(* IEC 61131-3 sources: daoli-st-library/DL_Process (part 13) *)

(* ---- FC_DL_GrateCoolerAirBalanceCalc.st ---- *)
(*
  Name: FC_DL_GrateCoolerAirBalanceCalc
  Category: DL_Process
  Version: 1.0.0
  Round: R91 / 2026-11-25
  开源溯源：clean-room 自研（族 水泥窑篦冷机与预热器，ST 开源生态实测 0 命中，无外部代码引入）
  功能：1) 篦冷机风量收支：把各风室冷却风量逐室求和得总冷却风量 fTotalAirNm3h，
           与窑头抽风（二次风 + 三次风 + 余风）合计 fDraftNm3h 做差，
           差值为正即「多余风量」（须经余风排放），差值为负即「亏缺风量」（抽风大于鼓风）。
        2) 不平衡率 fImbalancePct = |鼓风 − 抽风| / 鼓风 * 100，分母取鼓风侧（可测且恒正），
           方向固定不可交换；该值用于判断风量平衡是否在工艺允许带内。
        3) 平衡判据 fImbalancePct <= fBalMaxPct 输出 xBalanced，供上层选择「投自动调节」或「报警」。
  边界条件：1) 非有限值闸：九路实值入参先过 NOT(x > -DL_BIG AND x < DL_BIG)，同时拦 NaN 与 Inf，
           命中即闸断实值通路（全部输出强制 0.0），不得只置标志（R19）。
        2) 分母零闸：总冷却风量 |fTotalAirNm3h| <= DL_EPS 时不做除法，全部输出清零并判无效。
        3) 物理域闸：任一风室风量或抽风量为负即判无效（负风量属传感器反向或接线错误），
           不取绝对值掩盖符号错误；fBalMaxPct 须落在 (0.0, 100.0] 内，越域视为未组态。
        4) 判据取原始值（R24）：平衡判定使用钳制前的 _fImbalanceRawPct，不得先钳再判。
        5) 物理域钳制：不平衡率钳 0.0 ~ DL_PCT_HI；多余/亏缺风量钳 >= 0（两者互斥，只一支非零）。
        6) 单点赋值（R26）：多余与亏缺由同一差值按符号分支写入，先置 0 再按分支赋值一次，
           不在多处重复写同一变量；纯函数无状态，不做迟滞。
  量纲自证：fTotalAirNm3h / fDraftNm3h / fExcessNm3h / fDeficitNm3h 均为标态体积流量 [Nm3/h]，
           求和与求差两侧同量纲；
           fImbalancePct = |(Nm3/h) − (Nm3/h)| / (Nm3/h) * 100 = 无因次百分数 [%]，量纲合法。
  修订历史 Revision :
    2026-11-25  v1.0.0  R91 首版
*)

FUNCTION FC_DL_GrateCoolerAirBalanceCalc : BOOL
VAR_INPUT
    fChamber1Nm3h    : REAL;   // 1 风室冷却风量 [Nm3/h] / Chamber 1 cooling air flow [Nm3/h]
    fChamber2Nm3h    : REAL;   // 2 风室冷却风量 [Nm3/h] / Chamber 2 cooling air flow [Nm3/h]
    fChamber3Nm3h    : REAL;   // 3 风室冷却风量 [Nm3/h] / Chamber 3 cooling air flow [Nm3/h]
    fChamber4Nm3h    : REAL;   // 4 风室冷却风量 [Nm3/h] / Chamber 4 cooling air flow [Nm3/h]
    fChamber5Nm3h    : REAL;   // 5 风室冷却风量 [Nm3/h] / Chamber 5 cooling air flow [Nm3/h]
    fChamber6Nm3h    : REAL;   // 6 风室冷却风量 [Nm3/h] / Chamber 6 cooling air flow [Nm3/h]
    fDraftNm3h       : REAL;   // 窑头抽风合计（二次+三次+余风）[Nm3/h] / Total kiln-head draft [Nm3/h]
    fBalMaxPct       : REAL;   // 风量平衡允许不平衡率 [%] / Permitted imbalance ratio [%]
END_VAR
VAR_OUTPUT
    fTotalAirNm3h    : REAL;   // 各风室冷却风量合计 [Nm3/h] / Total cooling air flow [Nm3/h]
    fExcessNm3h      : REAL;   // 多余风量（鼓风大于抽风）[Nm3/h] / Excess air flow, blow over draft [Nm3/h]
    fDeficitNm3h     : REAL;   // 亏缺风量（抽风大于鼓风）[Nm3/h] / Deficit air flow, draft over blow [Nm3/h]
    fImbalancePct    : REAL;   // 风量不平衡率 [%] / Air balance imbalance ratio [%]
    xBalanced        : BOOL;   // 风量在允许带内 [bool] / Air balance within tolerance [bool]
    xValid           : BOOL;   // 计算有效标志 [bool] / Calculation valid flag [bool]
END_VAR
VAR
    _fDiffNm3h       : REAL;   // 鼓风减抽风的有符号差值 [Nm3/h] / Signed difference, blow minus draft [Nm3/h]
    _fImbalanceRawPct : REAL;  // 钳制前的不平衡率 [%] / Raw imbalance ratio before limiting [%]
END_VAR
VAR CONSTANT
    DL_EPS           : REAL := 1.0E-9;    // 数值零闸阈值 [-] / Numeric zero gate threshold [-]
    DL_BIG           : REAL := 1.0E12;    // 非有限值闸量级上限 [-] / Finiteness gate magnitude [-]
    DL_PCT           : REAL := 100.0;     // 百分比换算因子 [%] / Percent conversion factor [%]
    DL_PCT_HI        : REAL := 100.0;     // 不平衡率物理上限 [%] / Imbalance physical upper bound [%]
    DL_ZERO_NM3H     : REAL := 0.0;       // 风量零基准 [Nm3/h] / Zero flow reference [Nm3/h]
END_VAR

(* —— 段 1：非有限值闸（R19：闸断实值通路） —— *)
IF NOT (fChamber1Nm3h > -DL_BIG AND fChamber1Nm3h < DL_BIG)
   OR NOT (fChamber2Nm3h > -DL_BIG AND fChamber2Nm3h < DL_BIG)
   OR NOT (fChamber3Nm3h > -DL_BIG AND fChamber3Nm3h < DL_BIG)
   OR NOT (fChamber4Nm3h > -DL_BIG AND fChamber4Nm3h < DL_BIG)
   OR NOT (fChamber5Nm3h > -DL_BIG AND fChamber5Nm3h < DL_BIG)
   OR NOT (fChamber6Nm3h > -DL_BIG AND fChamber6Nm3h < DL_BIG)
   OR NOT (fDraftNm3h > -DL_BIG AND fDraftNm3h < DL_BIG)
   OR NOT (fBalMaxPct > -DL_BIG AND fBalMaxPct < DL_BIG) THEN
    fTotalAirNm3h := 0.0;                   // 输出强制 0.0，切断污染源 / Force zero, cut polluted path
    fExcessNm3h := 0.0;                     // 多余风量强制 0.0 / Excess forced to zero
    fDeficitNm3h := 0.0;                    // 亏缺风量强制 0.0 / Deficit forced to zero
    fImbalancePct := 0.0;                   // 不平衡率强制 0.0 / Imbalance forced to zero
    xBalanced := FALSE;                     // 失效侧不得报平衡 / Must not report balanced when invalid
    xValid := FALSE;                        // 有效位清零 / Validity cleared
    FC_DL_GrateCoolerAirBalanceCalc := FALSE;   // 返回码与有效位同源 / Return mirrors validity
    RETURN;                                 // 立即退出 / Immediate exit
END_IF

(* —— 段 2：风量求和（六室逐室相加，加法顺序不影响结果） —— *)
fTotalAirNm3h := fChamber1Nm3h + fChamber2Nm3h + fChamber3Nm3h
                 + fChamber4Nm3h + fChamber5Nm3h + fChamber6Nm3h;                  // 鼓风合计 [Nm3/h]
_fDiffNm3h := fTotalAirNm3h - fDraftNm3h;                                          // 鼓风 − 抽风 [Nm3/h]

(* —— 段 3：分母零闸（不平衡率的分母是鼓风合计） —— *)
IF ABS(fTotalAirNm3h) <= DL_EPS THEN
    fExcessNm3h := 0.0;                     // 无鼓风即无多余 / No blow, no excess
    fDeficitNm3h := 0.0;                    // 无鼓风即无亏缺 / No blow, no deficit
    fImbalancePct := 0.0;                   // 不平衡率不可算 / Imbalance not computable
    xBalanced := FALSE;                     // 判非平衡 / Not balanced
    xValid := FALSE;                        // 判无效 / Invalid
    FC_DL_GrateCoolerAirBalanceCalc := FALSE;   // 返回码同步 / Return synchronised
    RETURN;                                 // 提前退出 / Early exit
END_IF

_fImbalanceRawPct := ABS(_fDiffNm3h) / fTotalAirNm3h * DL_PCT;                    // 原始不平衡率 [%]

(* —— 段 4：判据（取原始值；单点 BOOL 聚合） —— *)
xValid := (fChamber1Nm3h >= DL_ZERO_NM3H)                                         // 各室风量不得为负
          AND (fChamber2Nm3h >= DL_ZERO_NM3H)
          AND (fChamber3Nm3h >= DL_ZERO_NM3H)
          AND (fChamber4Nm3h >= DL_ZERO_NM3H)
          AND (fChamber5Nm3h >= DL_ZERO_NM3H)
          AND (fChamber6Nm3h >= DL_ZERO_NM3H)
          AND (fDraftNm3h >= DL_ZERO_NM3H)                                        // 抽风量不得为负
          AND (fBalMaxPct > DL_EPS)                                               // 允许带必须为正
          AND (fBalMaxPct <= DL_PCT_HI);                                          // 允许带不得超过 100 %
xBalanced := xValid AND (_fImbalanceRawPct <= fBalMaxPct);                         // 在允许带内才算平衡

(* —— 段 5：多余/亏缺单点分支写入（互斥两支，各自只写一次，R26） —— *)
fExcessNm3h := 0.0;                                                               // 先置零，避免上拍残值
fDeficitNm3h := 0.0;                                                              // 先置零，避免上拍残值
IF _fDiffNm3h > DL_EPS THEN
    fExcessNm3h := _fDiffNm3h;                                                    // 鼓风大于抽风：多余 [Nm3/h]
ELSIF _fDiffNm3h < -DL_EPS THEN
    fDeficitNm3h := ABS(_fDiffNm3h);                                               // 抽风大于鼓风：亏缺 [Nm3/h]
END_IF

(* —— 段 6：输出单点写盘（不平衡率钳制到物理域） —— *)
fImbalancePct := LIMIT(0.0, _fImbalanceRawPct, DL_PCT_HI);                         // 不平衡率钳 0..100 [%]
FC_DL_GrateCoolerAirBalanceCalc := xValid;                                         // 返回码：TRUE = 计算可信

END_FUNCTION

(* ---- FC_DL_GrateCoolerBedResistanceCalc.st ---- *)
(*
  Name: FC_DL_GrateCoolerBedResistanceCalc
  Category: DL_Process
  Version: 1.0.0
  Round: R91 / 2026-11-25
  开源溯源：clean-room 自研（族 水泥窑篦冷机与预热器，ST 开源生态实测 0 命中，无外部代码引入）
  功能：1) 篦床料层阻力按「Ergun 型阻力式的粒度无关简化形」计算：压损正比于料层厚度、
           风量平方与料层堆积密度，反比于开孔率的三次方，
           即 dP = fK * H * rho * (Q/A_open)^2 / 2，A_open = A_total * phi，
           其中 fK 为综合阻力系数（含篦板结构与料层孔隙率经验项）。
        2) 输出三条派生量：料层压损 fBedDpKpa、按开孔率的等效穿孔风速 fOpenVelMs、
           以及压损相对上限的负荷率 fDpLoadPct（用于判断是否接近风机能力极限）。
        3) 压损上限 fDpMaxKpa 为设备许可值，超限只置 xValid=FALSE 并给出超限标志 xDpOver，
           数值本身钳到上限内输出，绝不把越限值伪装成合格值。
  边界条件：1) 非有限值闸：七路实值入参先过 NOT(x > -DL_BIG AND x < DL_BIG)，同时拦 NaN 与 Inf，
           命中即闸断实值通路（全部输出强制 0.0），不得只置标志（R19）。
        2) 分母零闸：料层厚度 fBedHeightM、篦床总面积 fGrateAreaM2 必须 > DL_EPS；
           开孔率 fOpenRatio 必须落在 (DL_PHI_EPS, 1.0] 内 —— 开孔率为 0 或大于 1 均属组态错误，
           直接判无效而非钳制，因为开孔率进三次方，钳制会严重扭曲结果。
        3) 判据取原始值（R24）：压损超限判定使用钳制前的 _fDpRawKpa，
           不得先把压损夹到上限再判是否越限（否则判据恒真）。
        4) 物理域钳制：压损钳 0.0 ~ fDpMaxKpa；穿孔风速钳 0.0 ~ DL_VEL_HI_MS；
           负荷率钳 0.0 ~ DL_LOAD_HI_PCT。
        5) 上限自身校验：fDpMaxKpa 必须 > DL_EPS，为负或零视为未组态，判无效。
        6) 纯函数无状态：不做去抖，堵塞判据的持续性与延时由下游监视 FB 承担。
  量纲自证：开孔面积 A_open = (m2)*(无因次) = m2；
           穿孔风速 = (m3/h)/(m2)/(s/h) = (m3/h)/(m2) * (h/s) = m/s；
           压损 = 无因次 * (m) * (kg/m3) * (m/s)^2 = (kg/m3)*(m2/s2)*(m) = kg/(m*s2) = Pa，
           再除 1000 得 kPa，量纲链自洽。
  修订历史 Revision :
    2026-11-25  v1.0.0  R91 首版
*)

FUNCTION FC_DL_GrateCoolerBedResistanceCalc : BOOL
VAR_INPUT
    fCoolingAirNm3h  : REAL;   // 该风室冷却风量 [Nm3/h] / Cooling air flow of the chamber [Nm3/h]
    fBedHeightM      : REAL;   // 篦床上料层厚度 [m] / Clinker bed height on the grate [m]
    fGrateAreaM2     : REAL;   // 该风室篦床有效面积 [m2] / Effective grate area of the chamber [m2]
    fOpenRatio       : REAL;   // 篦板开孔率（0~1 无因次）[-] / Grate open area ratio, dimensionless [-]
    fBulkDensityKgm3 : REAL;   // 料层堆积密度 [kg/m3] / Clinker bulk density [kg/m3]
    fResistCoef      : REAL;   // 综合阻力系数（含孔隙率经验项）[-] / Combined resistance coefficient [-]
    fDpMaxKpa        : REAL;   // 设备许可料层压损上限 [kPa] / Permitted bed pressure drop [kPa]
END_VAR
VAR_OUTPUT
    fBedDpKpa        : REAL;   // 料层压损 [kPa] / Clinker bed pressure drop [kPa]
    fOpenVelMs       : REAL;   // 篦板穿孔风速 [m/s] / Open-area jet velocity [m/s]
    fDpLoadPct       : REAL;   // 压损对上限的负荷率 [%] / Pressure drop load ratio [%]
    xDpOver          : BOOL;   // 压损超限标志（判定用原始值）[bool] / Pressure drop overrun flag [bool]
    xValid           : BOOL;   // 计算有效标志 [bool] / Calculation valid flag [bool]
END_VAR
VAR
    _fOpenAreaM2     : REAL;   // 篦板有效开孔面积 [m2] / Effective open area of the grate [m2]
    _fOpenVelRawMs   : REAL;   // 钳制前的穿孔风速 [m/s] / Raw open-area velocity [m/s]
    _fDpRawKpa       : REAL;   // 钳制前的原始料层压损 [kPa] / Raw bed pressure drop [kPa]
    _fLoadRawPct     : REAL;   // 钳制前的原始负荷率 [%] / Raw load ratio [%]
END_VAR
VAR CONSTANT
    DL_EPS           : REAL := 1.0E-9;    // 数值零闸阈值 [-] / Numeric zero gate threshold [-]
    DL_PHI_EPS       : REAL := 1.0E-6;    // 开孔率下限阈值 [-] / Open-ratio low gate threshold [-]
    DL_BIG           : REAL := 1.0E12;    // 非有限值闸量级上限 [-] / Finiteness gate magnitude [-]
    DL_SEC_PER_H     : REAL := 3600.0;    // 小时到秒的时基折算 [s/h] / Seconds per hour [s/h]
    DL_PA_PER_KPA    : REAL := 1000.0;    // 帕到千帕的折算 [Pa/kPa] / Pascals per kilopascal [Pa/kPa]
    DL_PHI_HI        : REAL := 1.0;       // 开孔率物理上限 [-] / Open-ratio physical upper bound [-]
    DL_VEL_HI_MS     : REAL := 100.0;     // 穿孔风速物理上限 [m/s] / Jet velocity upper bound [m/s]
    DL_PCT           : REAL := 100.0;     // 百分比换算因子 [%] / Percent conversion factor [%]
    DL_LOAD_HI_PCT   : REAL := 100.0;     // 负荷率物理上限 [%] / Load ratio upper bound [%]
END_VAR

(* —— 段 1：非有限值闸（R19：闸断实值通路） —— *)
IF NOT (fCoolingAirNm3h > -DL_BIG AND fCoolingAirNm3h < DL_BIG)
   OR NOT (fBedHeightM > -DL_BIG AND fBedHeightM < DL_BIG)
   OR NOT (fGrateAreaM2 > -DL_BIG AND fGrateAreaM2 < DL_BIG)
   OR NOT (fOpenRatio > -DL_BIG AND fOpenRatio < DL_BIG)
   OR NOT (fBulkDensityKgm3 > -DL_BIG AND fBulkDensityKgm3 < DL_BIG)
   OR NOT (fResistCoef > -DL_BIG AND fResistCoef < DL_BIG)
   OR NOT (fDpMaxKpa > -DL_BIG AND fDpMaxKpa < DL_BIG) THEN
    fBedDpKpa := 0.0;                       // 输出强制 0.0，切断污染源 / Force zero, cut polluted path
    fOpenVelMs := 0.0;                      // 风速同样强制 0.0 / Velocity forced to zero
    fDpLoadPct := 0.0;                      // 负荷率强制 0.0 / Load ratio forced to zero
    xDpOver := FALSE;                       // 超限位不得在失效时置真 / Overrun must stay false when invalid
    xValid := FALSE;                        // 有效位清零 / Validity cleared
    FC_DL_GrateCoolerBedResistanceCalc := FALSE;   // 返回码与有效位同源 / Return mirrors validity
    RETURN;                                 // 立即退出 / Immediate exit
END_IF

(* —— 段 2：几何与组态域闸（开孔率进三次方，越域一律判无效而非钳制） —— *)
IF (fGrateAreaM2 <= DL_EPS)                                       // 篦床面积不可为零
   OR (fBedHeightM <= DL_EPS)                                     // 料层厚度不可为零
   OR (fOpenRatio <= DL_PHI_EPS)                                  // 开孔率不可为零
   OR (fOpenRatio > DL_PHI_HI)                                    // 开孔率不得大于 1
   OR (fDpMaxKpa <= DL_EPS) THEN                                  // 压损上限必须已组态
    fBedDpKpa := 0.0;                       // 几何不可用即无压损 / No geometry, no drop
    fOpenVelMs := 0.0;                      // 风速不可算 / Velocity not computable
    fDpLoadPct := 0.0;                      // 负荷率不可算 / Load ratio not computable
    xDpOver := FALSE;                       // 失效侧超限位保持假 / Overrun stays false
    xValid := FALSE;                        // 判无效 / Invalid
    FC_DL_GrateCoolerBedResistanceCalc := FALSE;   // 返回码同步 / Return synchronised
    RETURN;                                 // 提前退出 / Early exit
END_IF

(* —— 段 3：主算式（不钳制，先出原始值供段 4 判据使用，R24） —— *)
_fOpenAreaM2 := fGrateAreaM2 * fOpenRatio;                                        // 有效开孔面积 [m2]
_fOpenVelRawMs := fCoolingAirNm3h / _fOpenAreaM2 / DL_SEC_PER_H;                  // 穿孔风速 [m/s]
_fDpRawKpa := fResistCoef * fBedHeightM * fBulkDensityKgm3
              * _fOpenVelRawMs * _fOpenVelRawMs / DL_PA_PER_KPA;                  // 动压式压损 [kPa]
_fLoadRawPct := _fDpRawKpa / fDpMaxKpa * DL_PCT;                                  // 原始负荷率 [%]

(* —— 段 4：判据（全部取原始值；单点 BOOL 聚合避免多处赋 FALSE 覆盖） —— *)
xDpOver := (_fDpRawKpa > fDpMaxKpa);                                              // 压损越上限
xValid := (fCoolingAirNm3h >= 0.0)                                                // 风量不得为负
          AND (fBedHeightM >= 0.0)                                                // 料层厚度不得为负
          AND (fBulkDensityKgm3 > 0.0)                                            // 堆积密度必须为正
          AND (fResistCoef > 0.0)                                                 // 阻力系数必须为正
          AND (_fOpenVelRawMs >= 0.0)                                             // 风速不得为负
          AND (_fDpRawKpa >= 0.0);                                                // 压损不得为负（负压损属符号错误）

(* —— 段 5：输出单点写盘（钳制到物理域内，判定结果已在段 4 定案） —— *)
fBedDpKpa := LIMIT(0.0, _fDpRawKpa, fDpMaxKpa);                                   // 压损钳 0..上限 [kPa]
fOpenVelMs := LIMIT(0.0, _fOpenVelRawMs, DL_VEL_HI_MS);                           // 风速钳 0..上限 [m/s]
fDpLoadPct := LIMIT(0.0, _fLoadRawPct, DL_LOAD_HI_PCT);                           // 负荷率钳 0..100 [%]
FC_DL_GrateCoolerBedResistanceCalc := xValid;                                     // 返回码：TRUE = 计算可信

END_FUNCTION

(* ---- FC_DL_GrateCoolerClinkerTempCalc.st ---- *)
(*
  Name: FC_DL_GrateCoolerClinkerTempCalc
  Category: DL_Process
  Version: 1.0.0
  Round: R91 / 2026-11-25
  开源溯源：clean-room 自研（族 水泥窑篦冷机与预热器，ST 开源生态实测 0 命中，无外部代码引入）
  功能：1) 出篦冷机熟料温度按「熟料放热 = 空气吸热」的稳态能量平衡求解：
           熟料放热 = m_cli * cp_cli * (T_in − T_out)，空气吸热 = m_cli * ratio * cp_air * (T_airOut − T_airIn)，
           两式相等并引入换热效率 eff 后反解出口温度：
           T_out = T_in − eff * ratio * (cp_air / cp_cli) * (T_airOut − T_airIn)。
        2) 输出熟料降温幅度 fCoolDropK，即 T_in − T_out，用于判断冷却能力是否达标。
        3) 温度下限保护：反解结果不得低于 DL_TEMP_LO（环境温度下限），低于即判无效，
           因为能量平衡模型在该区间外已不成立（潜热与辐射项未建模）。
  边界条件：1) 非有限值闸：七路实值入参先过 NOT(x > -DL_BIG AND x < DL_BIG)，同时拦 NaN 与 Inf，
           命中即闸断实值通路（全部输出强制 0.0），不得只置标志（R19）。
        2) 分母零闸：熟料比热 fClinkerCpKjKgK 与风料比 fAirClinkerRatio 均须 > DL_EPS，
           否则反解式分母为零、结果发散，直接判无效。
        3) 参数域闸：换热效率 fEffRatio 必须落在 (0.0, 1.0] 内（效率大于 1 违反热力学第一定律），
           越域视为组态错误判无效，不钳制（钳制会把非法组态伪装成合法）。
        4) 温差方向闸：空气出口温度必须高于空气入口温度，否则无吸热过程，判无效。
        5) 温度下限：反解出口温度 < DL_TEMP_LO 判无效；上限 DL_TEMP_HI 越限判无效。
        6) 判据取原始值（R24）：温度越域判定使用原始反解值 _fOutRawC，钳制只作用于输出量。
  量纲自证：ratio 为风料质量比 [kg/kg] 无因次；cp_air / cp_cli = (kJ/(kg*K))/(kJ/(kg*K)) 无因次；
           eff 无因次；故 eff*ratio*(cp_air/cp_cli)*(T_airOut−T_airIn) 的量纲为 (K)，
           与 T_in [degC] 相减合法（温差以 K 计、绝对温度以 degC 计，差值同尺度）。
  修订历史 Revision :
    2026-11-25  v1.0.0  R91 首版
*)

FUNCTION FC_DL_GrateCoolerClinkerTempCalc : BOOL
VAR_INPUT
    fClinkerInC      : REAL;   // 入篦冷机熟料温度 [degC] / Clinker inlet temperature [degC]
    fAirInC          : REAL;   // 冷却风入口温度（环境）[degC] / Cooling air inlet temperature [degC]
    fAirOutC         : REAL;   // 冷却风出口温度（窑头抽风）[degC] / Cooling air outlet temperature [degC]
    fAirClinkerRatio : REAL;   // 风料质量比 [kg/kg] / Air to clinker mass ratio [kg/kg]
    fAirCpKjKgK      : REAL;   // 空气定压比热 [kJ/(kg*K)] / Air specific heat at constant pressure [kJ/(kg*K)]
    fClinkerCpKjKgK  : REAL;   // 熟料比热 [kJ/(kg*K)] / Clinker specific heat [kJ/(kg*K)]
    fEffRatio        : REAL;   // 篦床换热效率（0~1 无因次）[-] / Grate heat exchange efficiency, dimensionless [-]
END_VAR
VAR_OUTPUT
    fClinkerOutC     : REAL;   // 出篦冷机熟料温度 [degC] / Clinker outlet temperature [degC]
    fCoolDropK       : REAL;   // 熟料降温幅度 [K] / Clinker temperature drop [K]
    xTempLow         : BOOL;   // 出口温度低于下限标志 [bool] / Outlet below lower bound flag [bool]
    xValid           : BOOL;   // 计算有效标志 [bool] / Calculation valid flag [bool]
END_VAR
VAR
    _fCpRatio        : REAL;   // 空气与熟料比热之比 [-] / Ratio of air to clinker specific heat [-]
    _fAirDeltaK      : REAL;   // 空气温升 [K] / Air temperature rise [K]
    _fOutRawC        : REAL;   // 钳制前的原始出口温度 [degC] / Raw outlet temperature before limiting [degC]
    _fDropRawK       : REAL;   // 钳制前的原始降温幅度 [K] / Raw temperature drop before limiting [K]
END_VAR
VAR CONSTANT
    DL_EPS           : REAL := 1.0E-9;    // 数值零闸阈值 [-] / Numeric zero gate threshold [-]
    DL_BIG           : REAL := 1.0E12;    // 非有限值闸量级上限 [-] / Finiteness gate magnitude [-]
    DL_TEMP_LO       : REAL := -50.0;     // 熟料出口温度物理下限 [degC] / Clinker outlet lower bound [degC]
    DL_TEMP_HI       : REAL := 400.0;     // 熟料出口温度物理上限 [degC] / Clinker outlet upper bound [degC]
    DL_EFF_HI        : REAL := 1.0;       // 换热效率物理上限（热力学第一定律）[-] / Efficiency upper bound [-]
    DL_ZERO_K        : REAL := 0.0;       // 温差零基准 [K] / Zero temperature-difference reference [K]
END_VAR

(* —— 段 1：非有限值闸（R19：闸断实值通路） —— *)
IF NOT (fClinkerInC > -DL_BIG AND fClinkerInC < DL_BIG)
   OR NOT (fAirInC > -DL_BIG AND fAirInC < DL_BIG)
   OR NOT (fAirOutC > -DL_BIG AND fAirOutC < DL_BIG)
   OR NOT (fAirClinkerRatio > -DL_BIG AND fAirClinkerRatio < DL_BIG)
   OR NOT (fAirCpKjKgK > -DL_BIG AND fAirCpKjKgK < DL_BIG)
   OR NOT (fClinkerCpKjKgK > -DL_BIG AND fClinkerCpKjKgK < DL_BIG)
   OR NOT (fEffRatio > -DL_BIG AND fEffRatio < DL_BIG) THEN
    fClinkerOutC := 0.0;                    // 输出强制 0.0，切断污染源 / Force zero, cut polluted path
    fCoolDropK := 0.0;                      // 降温幅度强制 0.0 / Drop forced to zero
    xTempLow := FALSE;                      // 失效侧不得报低温 / Must not report low temp when invalid
    xValid := FALSE;                        // 有效位清零 / Validity cleared
    FC_DL_GrateCoolerClinkerTempCalc := FALSE;   // 返回码与有效位同源 / Return mirrors validity
    RETURN;                                 // 立即退出 / Immediate exit
END_IF

(* —— 段 2：分母零闸与参数域闸（比热、风料比为零则反解发散） —— *)
IF (fClinkerCpKjKgK <= DL_EPS)                                    // 熟料比热不可为零
   OR (fAirClinkerRatio <= DL_EPS)                                // 风料比不可为零
   OR (fAirCpKjKgK <= DL_EPS)                                     // 空气比热不可为零
   OR (fEffRatio <= DL_EPS)                                       // 换热效率不可为零
   OR (fEffRatio > DL_EFF_HI) THEN                                // 换热效率不得大于 1（热力学第一定律）
    fClinkerOutC := 0.0;                    // 参数不可用即无出口温度 / No parameter, no outlet temperature
    fCoolDropK := 0.0;                      // 降温幅度不可算 / Drop not computable
    xTempLow := FALSE;                      // 失效侧低温位保持假 / Low-temp flag stays false
    xValid := FALSE;                        // 判无效 / Invalid
    FC_DL_GrateCoolerClinkerTempCalc := FALSE;   // 返回码同步 / Return synchronised
    RETURN;                                 // 提前退出 / Early exit
END_IF

(* —— 段 3：主算式（不钳制，先出原始值供段 4 判据使用，R24） —— *)
_fCpRatio := fAirCpKjKgK / fClinkerCpKjKgK;                                       // 比热之比 [-]
_fAirDeltaK := fAirOutC - fAirInC;                                                // 空气温升 [K]
_fOutRawC := fClinkerInC - fEffRatio * fAirClinkerRatio * _fCpRatio * _fAirDeltaK; // 出口温度反解 [degC]
_fDropRawK := fClinkerInC - _fOutRawC;                                            // 降温幅度 [K]

(* —— 段 4：判据（取原始值；单点 BOOL 聚合避免多处赋 FALSE 覆盖） —— *)
xTempLow := (_fOutRawC < DL_TEMP_LO);                                             // 出口低于物理下限
xValid := (_fAirDeltaK > DL_ZERO_K)                                               // 空气必须吸热（出口高于入口）
          AND (_fOutRawC >= DL_TEMP_LO)                                           // 不跌破物理下限
          AND (_fOutRawC <= DL_TEMP_HI)                                           // 不超出物理上限
          AND (_fDropRawK >= DL_ZERO_K)                                           // 降温幅度不得为负（方向固定）
          AND (fClinkerInC > DL_TEMP_LO);                                         // 入口温度本身须在物理域内

(* —— 段 5：输出单点写盘（钳制到物理域内，判定结果已在段 4 定案） —— *)
fClinkerOutC := LIMIT(DL_TEMP_LO, _fOutRawC, DL_TEMP_HI);                          // 出口温度钳物理域 [degC]
fCoolDropK := MAX(DL_ZERO_K, _fDropRawK);                                          // 降温幅度钳 >= 0 [K]
FC_DL_GrateCoolerClinkerTempCalc := xValid;                                        // 返回码：TRUE = 计算可信

END_FUNCTION

(* ---- FC_DL_GrateCoolerHeatRecoveryCalc.st ---- *)
(*
  Name: FC_DL_GrateCoolerHeatRecoveryCalc
  Category: DL_Process
  Version: 1.0.0
  Round: R91 / 2026-11-25
  开源溯源：clean-room 自研（族 水泥窑篦冷机与预热器，ST 开源生态实测 0 命中，无外部代码引入）
  功能：1) 回收热量取「二次风显热 + 三次风显热」，两者均以环境温度为基准，风侧按定压比热折算，
           即 fRecoveredHeatKw = (V2*cp*(T2-Tamb) + V3*cp*(T3-Tamb)) / 3600，单位 kW，
           3600 为 kJ/h 到 kW 的时基折算系数。
        2) 熟料可供显热取「熟料量 × 熟料比热 × (入篦床温度 − 出篦床温度)」，
           即 fClinkerHeatKw = m*1000*cpCli*(Tin-Tout) / 3600，单位 kW，
           1000 为 t 到 kg 的质量折算系数；该项是回收率的物理分母（可供热上限）。
        3) 热回收率 fRecoveryPct = 回收热量 / 熟料可供显热 * 100，钳制 0.0 ~ 100.0 %，
           回收率超过 100 % 在物理上不可能，判为测量链路故障而非效率优异。
  边界条件：1) 非有限值闸：九路实值入参先过 NOT(x > -DL_BIG AND x < DL_BIG)，该式同时拦 NaN 与 Inf，
           命中即闸断实值通路（全部输出强制 0.0），不得只置 xValid 而把 NaN 传给下游（R19）。
        2) 分母零闸：风侧比热 fAirCpKjNm3K 与熟料比热 fClinkerCp 均须 > DL_EPS，
           熟料可供显热 |fClinkerHeatKw| > DL_EPS 才允许做除法，否则判无效并清零。
        3) 判据取原始值（R24）：回收率越限判定使用 LIMIT 之前的原始值 _fRecoveryRawPct，
           不得先把回收率夹到 0~100 再判超域（否则判据恒真，域闸静默失效）。
        4) 物理域钳制：回收率钳 0.0 ~ 100.0 %；两路风量与熟料量不得为负（负值即传感器反向，判无效）。
        5) 温度方向校验：二次/三次风温低于环境温度、或熟料出口温度高于入口温度，均属非冷却工况，
           判无效而不取绝对值掩盖符号错误。
        6) 纯函数无状态：本件不做迟滞与去抖，滤波与报警延时由下游监视 FB 承担。
  量纲自证：fRecoveredHeatKw = (Nm3/h)*(kJ/(Nm3*K))*(K) / (s/h) = (kJ/h)/(s/h) = kJ/s = kW；
           fClinkerHeatKw   = (t/h)*(kg/t)*(kJ/(kg*K))*(K) / (s/h) = (kJ/h)/(s/h) = kW；
           fRecoveryPct     = (kW)/(kW)*100 = 无因次百分数 [%]，比量两侧同量纲，量纲关系合法。
  修订历史 Revision :
    2026-11-25  v1.0.0  R91 首版
*)

FUNCTION FC_DL_GrateCoolerHeatRecoveryCalc : BOOL
VAR_INPUT
    fSecAirNm3h      : REAL;   // 二次风标态体积流量 [Nm3/h] / Secondary air normal flow [Nm3/h]
    fTerAirNm3h      : REAL;   // 三次风标态体积流量 [Nm3/h] / Tertiary air normal flow [Nm3/h]
    fSecAirTempC     : REAL;   // 二次风温度 [degC] / Secondary air temperature [degC]
    fTerAirTempC     : REAL;   // 三次风温度 [degC] / Tertiary air temperature [degC]
    fAmbientC        : REAL;   // 环境基准温度 [degC] / Ambient reference temperature [degC]
    fClinkerTph      : REAL;   // 熟料产量 [t/h] / Clinker production rate [t/h]
    fClinkerInC      : REAL;   // 入篦床熟料温度 [degC] / Clinker inlet temperature [degC]
    fClinkerOutC     : REAL;   // 出篦床熟料温度 [degC] / Clinker outlet temperature [degC]
    fAirCpKjNm3K     : REAL;   // 风侧定压比热 [kJ/(Nm3*K)] / Air specific heat at constant pressure [kJ/(Nm3*K)]
    fClinkerCpKjKgK  : REAL;   // 熟料比热 [kJ/(kg*K)] / Clinker specific heat [kJ/(kg*K)]
END_VAR
VAR_OUTPUT
    fRecoveredHeatKw : REAL;   // 二次+三次风回收热量 [kW] / Recovered heat by secondary and tertiary air [kW]
    fClinkerHeatKw   : REAL;   // 熟料可供显热 [kW] / Clinker available sensible heat [kW]
    fRecoveryPct     : REAL;   // 热回收率 [%] / Heat recovery ratio [%]
    xValid           : BOOL;   // 计算有效标志 [bool] / Calculation valid flag [bool]
END_VAR
VAR
    _fSecHeatKjh     : REAL;   // 二次风显热 [kJ/h] / Secondary air sensible heat [kJ/h]
    _fTerHeatKjh     : REAL;   // 三次风显热 [kJ/h] / Tertiary air sensible heat [kJ/h]
    _fRecoveredKjh   : REAL;   // 回收热量合计（钳制前）[kJ/h] / Total recovered heat before limiting [kJ/h]
    _fClinkerKjh     : REAL;   // 熟料可供显热（钳制前）[kJ/h] / Clinker sensible heat before limiting [kJ/h]
    _fRecoveryRawPct : REAL;   // 钳制前的原始回收率 [%] / Raw recovery before limiting [%]
END_VAR
VAR CONSTANT
    DL_EPS           : REAL := 1.0E-9;    // 数值零闸阈值 [-] / Numeric zero gate threshold [-]
    DL_BIG           : REAL := 1.0E12;    // 非有限值闸量级上限 [-] / Finiteness gate magnitude [-]
    DL_SEC_PER_H     : REAL := 3600.0;    // 小时到秒的时基折算 [s/h] / Seconds per hour [s/h]
    DL_KG_PER_T      : REAL := 1000.0;    // 吨到千克的质量折算 [kg/t] / Kilograms per tonne [kg/t]
    DL_PCT           : REAL := 100.0;     // 百分比换算因子 [%] / Percent conversion factor [%]
    DL_REC_LO_PCT    : REAL := 0.0;       // 回收率物理域下限 [%] / Recovery physical domain low [%]
    DL_REC_HI_PCT    : REAL := 100.0;     // 回收率物理域上限 [%] / Recovery physical domain high [%]
END_VAR

(* —— 段 1：非有限值闸（R19：闸断实值通路，NaN/Inf 一律不得流到输出） —— *)
IF NOT (fSecAirNm3h > -DL_BIG AND fSecAirNm3h < DL_BIG)
   OR NOT (fTerAirNm3h > -DL_BIG AND fTerAirNm3h < DL_BIG)
   OR NOT (fSecAirTempC > -DL_BIG AND fSecAirTempC < DL_BIG)
   OR NOT (fTerAirTempC > -DL_BIG AND fTerAirTempC < DL_BIG)
   OR NOT (fAmbientC > -DL_BIG AND fAmbientC < DL_BIG)
   OR NOT (fClinkerTph > -DL_BIG AND fClinkerTph < DL_BIG)
   OR NOT (fClinkerInC > -DL_BIG AND fClinkerInC < DL_BIG)
   OR NOT (fClinkerOutC > -DL_BIG AND fClinkerOutC < DL_BIG)
   OR NOT (fAirCpKjNm3K > -DL_BIG AND fAirCpKjNm3K < DL_BIG)
   OR NOT (fClinkerCpKjKgK > -DL_BIG AND fClinkerCpKjKgK < DL_BIG) THEN
    fRecoveredHeatKw := 0.0;                // 输出强制 0.0，切断污染源 / Force zero, cut polluted path
    fClinkerHeatKw := 0.0;                  // 熟料显热同样强制 0.0 / Clinker heat forced to zero
    fRecoveryPct := 0.0;                    // 回收率强制 0.0 / Recovery forced to zero
    xValid := FALSE;                        // 有效位清零 / Validity cleared
    FC_DL_GrateCoolerHeatRecoveryCalc := FALSE;   // 返回码与有效位同源 / Return mirrors validity
    RETURN;                                 // 立即退出 / Immediate exit
END_IF

(* —— 段 2：比热零闸（R4：除法前先过零闸，且闸的是分母本身） —— *)
IF ABS(fAirCpKjNm3K) <= DL_EPS OR ABS(fClinkerCpKjKgK) <= DL_EPS THEN
    fRecoveredHeatKw := 0.0;                // 比热缺失即无法折算 / No specific heat, no conversion
    fClinkerHeatKw := 0.0;                  // 熟料显热不可算 / Clinker heat not computable
    fRecoveryPct := 0.0;                    // 回收率不可算 / Recovery not computable
    xValid := FALSE;                        // 判无效 / Invalid
    FC_DL_GrateCoolerHeatRecoveryCalc := FALSE;   // 返回码同步 / Return synchronised
    RETURN;                                 // 提前退出 / Early exit
END_IF

(* —— 段 3：主算式（不做任何钳制，先出原始值供段 4 判据使用，R24） —— *)
_fSecHeatKjh := fSecAirNm3h * fAirCpKjNm3K * (fSecAirTempC - fAmbientC);          // 二次风显热 [kJ/h]
_fTerHeatKjh := fTerAirNm3h * fAirCpKjNm3K * (fTerAirTempC - fAmbientC);          // 三次风显热 [kJ/h]
_fRecoveredKjh := _fSecHeatKjh + _fTerHeatKjh;                                    // 回收热量合计 [kJ/h]
_fClinkerKjh := fClinkerTph * DL_KG_PER_T * fClinkerCpKjKgK
                * (fClinkerInC - fClinkerOutC);                                   // 熟料可供显热 [kJ/h]

(* —— 段 4：分母零闸（熟料可供显热为回收率的分母） —— *)
IF ABS(_fClinkerKjh) <= DL_EPS THEN
    fRecoveredHeatKw := 0.0;                // 无可供热即无回收率 / No source heat, no recovery
    fClinkerHeatKw := 0.0;                  // 分母侧同步清零 / Denominator side zeroed
    fRecoveryPct := 0.0;                    // 回收率清零 / Recovery zeroed
    xValid := FALSE;                        // 判无效 / Invalid
    FC_DL_GrateCoolerHeatRecoveryCalc := FALSE;   // 返回码同步 / Return synchronised
    RETURN;                                 // 提前退出 / Early exit
END_IF

_fRecoveryRawPct := _fRecoveredKjh / _fClinkerKjh * DL_PCT;                       // 原始回收率 [%]

(* —— 段 5：物理域与符号校验（判据全部取原始值，单点 BOOL 聚合避免多处赋 FALSE 覆盖） —— *)
xValid := (fSecAirNm3h >= 0.0)                                        // 二次风量不得为负
          AND (fTerAirNm3h >= 0.0)                                    // 三次风量不得为负
          AND (fClinkerTph >= 0.0)                                    // 熟料量不得为负
          AND (_fRecoveredKjh >= 0.0)                                 // 风温低于环境温度属非回收工况
          AND (_fClinkerKjh > 0.0)                                    // 熟料出口必须低于入口
          AND (_fRecoveryRawPct >= DL_REC_LO_PCT)                     // 不低于物理域下限
          AND (_fRecoveryRawPct <= DL_REC_HI_PCT);                    // 不高于物理域上限（>100 % 物理不可能）

(* —— 段 6：输出单点写盘（数值钳制到物理域内，有效位已在段 5 定案） —— *)
fRecoveredHeatKw := _fRecoveredKjh / DL_SEC_PER_H;                                        // 折算为 kW
fClinkerHeatKw := _fClinkerKjh / DL_SEC_PER_H;                                            // 折算为 kW
fRecoveryPct := LIMIT(DL_REC_LO_PCT, _fRecoveryRawPct, DL_REC_HI_PCT);                    // 回收率钳 0..100 [%]
FC_DL_GrateCoolerHeatRecoveryCalc := xValid;                                              // 返回码：TRUE = 计算可信

END_FUNCTION

(* ---- FC_DL_GreenSandCompactabilityCalc.st ---- *)
(*
 * FC_DL_GreenSandCompactabilityCalc | C1 | DL_Process
 * 功能：由含水量反算紧实率并判定是否落在工艺带       单位：水分 [%]、紧实率 [%]、系数 [%/%、1]
 * 工况边界：w = a + b×CB 的反解 CB = (w−a)/b，b 须 >0（本件强制 b≠0，否则判 9714）；工艺带 30~45 %（含端点，浮点比较用容差）；a、b 与水分须有限
 * 代数值回代：w=3.0 %、a=1.2、b=0.04 → CB=(3.0−1.2)/0.04=45 %，落在 30~45 → xInRange=TRUE（与 spec 回代行一致）
 * 开源溯源：clean-room 自研，未复制任何第三方代码（无外部来源）
 *)
FUNCTION FC_DL_GreenSandCompactabilityCalc : BOOL
VAR_INPUT
    rMoisturePct : REAL := 3.0;      // 型砂含水量 | green sand moisture [%]
    rA           : REAL := 1.2;      // 经验式截距 | empirical intercept [%]
    rB           : REAL := 0.04;     // 经验式斜率 | empirical slope [%/%]
END_VAR
VAR_OUTPUT
    rCompactabilityPct : REAL;       // 紧实率 | compactability [%]
    xInRange           : BOOL;       // 落在工艺带 30~45 | inside the process band 30 to 45
    xValid             : BOOL;       // 输出有效 | outputs valid
    nFaultCode         : INT;        // 0=无 / 9714=斜率或水分非法 | 0 none, 9714 illegal slope or moisture
END_VAR
VAR
    xFinW : BOOL;                    // 水分有限性 | moisture is finite
    xFinA : BOOL;                    // 截距有限性 | intercept is finite
    xFinB : BOOL;                    // 斜率有限性 | slope is finite
END_VAR
VAR CONSTANT
    DL_GSC_LO  : REAL := 30.0;       // 工艺带下限 | process band lower bound [%]
    DL_GSC_HI  : REAL := 45.0;       // 工艺带上限 | process band upper bound [%]
    DL_GSC_EPS : REAL := 1.0E-6;     // 浮点比较容差 | floating comparison tolerance [%]
    DL_GSC_BMIN: REAL := 1.0E-9;     // 斜率下限（防零除）| slope lower bound guarding the division [%/%]
END_VAR

// 段1｜非有限闸（R19）
xFinW := (rMoisturePct = rMoisturePct) AND ((rMoisturePct - rMoisturePct) = 0.0);
xFinA := (rA = rA) AND ((rA - rA) = 0.0);
xFinB := (rB = rB) AND ((rB - rB) = 0.0);
IF (NOT xFinW) OR (NOT xFinA) OR (NOT xFinB) THEN
    rCompactabilityPct := 0.0;       // 安全值：紧实率 0 | safe value, zero compactability
    xInRange := FALSE;
    xValid := FALSE;
    nFaultCode := 9714;
    FC_DL_GreenSandCompactabilityCalc := FALSE;
    RETURN;
END_IF

// 段2｜域闸：斜率入分母必须为正，水分不得为负
IF (rB <= DL_GSC_BMIN) OR (rMoisturePct < 0.0) THEN
    rCompactabilityPct := 0.0;
    xInRange := FALSE;
    xValid := FALSE;
    nFaultCode := 9714;
    FC_DL_GreenSandCompactabilityCalc := FALSE;
    RETURN;
END_IF

// 段3｜算法：CB = (w − a)/b
rCompactabilityPct := (rMoisturePct - rA) / rB;

// 段4｜工艺带判定（判据与出口同源于原始水分推算值）
xInRange := (rCompactabilityPct >= (DL_GSC_LO - DL_GSC_EPS))
             AND (rCompactabilityPct <= (DL_GSC_HI + DL_GSC_EPS));
nFaultCode := 0;
xValid := TRUE;
FC_DL_GreenSandCompactabilityCalc := TRUE;
END_FUNCTION

(* ---- FC_DL_GreenSandMoistureTargetCalc.st ---- *)
(*
 * FC_DL_GreenSandMoistureTargetCalc | C2 | DL_Process
 * 功能：由紧实率反算湿型砂水分目标（线性经验式）       单位：紧实率 [%]、水分 [%]、系数 [%/%、1]
 * 工况边界：经验式 w = a + b×CB，a=1.2 %、b=0.04 %/%（spec 采纳值，回代 38 → 2.72 %，落在湿型砂 2.5~3.5 % 合理区间）；紧实率按物理域钳位 [20,60] %，越界置信息位且判据取自未钳位原值；系数 b 须 >0
 * 代数值回代：CB=38 %、a=1.2、b=0.04 → w=1.2+0.04×38=2.72 %（与 spec 采纳回代值一致）
 * 系数修正说明：spec 初版给 a=0.55 / b=0.0525，回代 38 得 2.545 % 偏离湿型砂常规区间，spec 已明确改用 a=1.2 / b=0.04，本件按采纳值实现
 * 开源溯源：clean-room 自研，未复制任何第三方代码（无外部来源）
 *)
FUNCTION FC_DL_GreenSandMoistureTargetCalc : BOOL
VAR_INPUT
    rCompactabilityPct : REAL := 38.0;  // 紧实率 | compactability [%]
    rA                 : REAL := 1.2;   // 经验式截距 | empirical intercept [%]
    rB                 : REAL := 0.04;  // 经验式斜率 | empirical slope [%/%]
END_VAR
VAR_OUTPUT
    rTargetMoisturePct : REAL;          // 目标水分 | target moisture [%]
    rCbUsed            : REAL;          // 实际参与计算的紧实率（已钳位）| compactability actually used, clamped [%]
    xClamped           : BOOL;          // 紧实率越界被钳位（信息级）| compactability clamped, informational
    xValid             : BOOL;          // 输出有效 | outputs valid
END_VAR
VAR
    xFinCb : BOOL;                      // 紧实率有限性 | compactability is finite
    xFinA  : BOOL;                      // 截距有限性 | intercept is finite
    xFinB  : BOOL;                      // 斜率有限性 | slope is finite
END_VAR
VAR CONSTANT
    DL_GSM_CB_LO : REAL := 20.0;        // 紧实率物理下限 | compactability lower bound [%]
    DL_GSM_CB_HI : REAL := 60.0;        // 紧实率物理上限 | compactability upper bound [%]
END_VAR

// 段1｜非有限闸（R19）
xFinCb := (rCompactabilityPct = rCompactabilityPct) AND ((rCompactabilityPct - rCompactabilityPct) = 0.0);
xFinA := (rA = rA) AND ((rA - rA) = 0.0);
xFinB := (rB = rB) AND ((rB - rB) = 0.0);
IF (NOT xFinCb) OR (NOT xFinA) OR (NOT xFinB) THEN
    rTargetMoisturePct := 0.0;          // 安全值：目标水分 0 | safe value, zero target
    rCbUsed := 0.0;
    xClamped := FALSE;
    xValid := FALSE;
    FC_DL_GreenSandMoistureTargetCalc := FALSE;
    RETURN;
END_IF

// 段2｜域闸：斜率必须为正（经验式单调增，否则反算无意义）
IF rB <= 0.0 THEN
    rTargetMoisturePct := 0.0;
    rCbUsed := 0.0;
    xClamped := FALSE;
    xValid := FALSE;
    FC_DL_GreenSandMoistureTargetCalc := FALSE;
    RETURN;
END_IF

// 段3｜域钳位：越界标志取自未钳位原值（R24）
IF rCompactabilityPct < DL_GSM_CB_LO THEN
    xClamped := TRUE;
    rCbUsed := DL_GSM_CB_LO;
ELSIF rCompactabilityPct > DL_GSM_CB_HI THEN
    xClamped := TRUE;
    rCbUsed := DL_GSM_CB_HI;
ELSE
    xClamped := FALSE;
    rCbUsed := rCompactabilityPct;
END_IF

// 段4｜算法：w = a + b×CB
rTargetMoisturePct := rA + rB * rCbUsed;
xValid := TRUE;
FC_DL_GreenSandMoistureTargetCalc := TRUE;
END_FUNCTION

(* ---- FC_DL_GreenStrengthIndexCalc.st ---- *)
(*
  Component : FC_DL_GreenStrengthIndexCalc
  Category  : DL_Process
  Type      : FC
  Complexity: C2
  VERSION   : v1.0.0
  功能      : 生坯强度指数核算：按压制成型压力、润滑剂含量与生坯密度算无量纲强度指数，并与安全阈值比较给出脱模安全判定。
  开源溯源  : 道莅原创 clean-room 自研（无外部代码引用）｜License: MIT
  边界条件  : ① 参考密度与安全阈值须 > 1e-9，压制压力须非负，润滑剂含量须在 0~5 % 内，否则返回哨兵 -1；
              ② 压力项取开方（压力对强度是次线性贡献），开方前已钳位非负；
              ③ 润滑剂含量越高生坯强度越低，折算系数下限钳位 0.3。
*)
FUNCTION FC_DL_GreenStrengthIndexCalc : REAL
VAR_INPUT
    fPressMPa    : REAL;   (* 压制压力 [MPa] Compaction pressure *)
    fLubePct     : REAL;   (* 润滑剂含量 [%] Lubricant content *)
    fGreenDens   : REAL;   (* 生坯密度 [g/cm³] Green density *)
    fDensRef     : REAL;   (* 参考密度（工艺目标） [g/cm³] Reference density *)
    fSafeIdx     : REAL;   (* 脱模安全指数阈值 [-] Safe ejection index threshold *)
END_VAR
VAR_OUTPUT
    fStrengthIdx : REAL;  (* 生坯强度指数 [-] Green strength index *)
    fLubeFactor  : REAL;  (* 润滑剂折减因子 [-] Lubricant reduction factor *)
    xEjectSafe   : BOOL;  (* 脱模安全标志 [-] Safe ejection flag *)
    xValid       : BOOL;  (* 计算有效性标志 [-] Calculation valid flag *)
END_VAR
VAR CONSTANT
    DL_EPS      : REAL := 1.0E-9;   (* 除零判定容差 [无量纲] Divide-by-zero tolerance *)
    DL_PCT_BASE : REAL := 100.0;    (* 百分比基准 [%] Percent base *)
    DL_GAIN     : REAL := 3.0;      (* 压力项标定增益 [-] Pressure term gain *)
    DL_LUBE_K   : REAL := 0.9;      (* 润滑剂折减系数 [-] Lubricant reduction coefficient *)
    DL_LUBE_MAX : REAL := 5.0;      (* 润滑剂含量上限 [%] Lubricant upper bound *)
    DL_LF_MIN   : REAL := 0.3;      (* 润滑剂因子下限 [-] Lubricant factor floor *)
    DL_ZERO     : REAL := 0.0;      (* 零常量 [无量纲] Zero constant *)
END_VAR
VAR
    fPressPos : REAL;   (* 非负压制压力 [MPa] Non-negative pressure *)
END_VAR
(* 出口预置：四出口统一预置 *)
fStrengthIdx := 0.0; fLubeFactor := 1.0; xEjectSafe := FALSE; xValid := FALSE;
(* 非有限拦截：自反判 NaN，自身差值判 Inf *)
IF (fPressMPa <> fPressMPa) OR ((fPressMPa - fPressMPa) <> 0.0)
   OR (fLubePct <> fLubePct) OR ((fLubePct - fLubePct) <> 0.0)
   OR (fGreenDens <> fGreenDens) OR ((fGreenDens - fGreenDens) <> 0.0)
   OR (fDensRef <> fDensRef) OR ((fDensRef - fDensRef) <> 0.0)
   OR (fSafeIdx <> fSafeIdx) OR ((fSafeIdx - fSafeIdx) <> 0.0) THEN
    FC_DL_GreenStrengthIndexCalc := -1.0;  (* 哨兵 -1：输入非有限 / Sentinel -1 non-finite *)
    RETURN;
END_IF
(* 组态域闸：参考密度与安全阈值为比例基，润滑剂含量与压力取可表区间 *)
IF (fDensRef <= DL_EPS) OR (fSafeIdx <= DL_EPS) OR (fPressMPa < DL_ZERO)
   OR (fLubePct < DL_ZERO) OR (fLubePct > DL_LUBE_MAX) OR (fGreenDens < DL_ZERO) THEN
    FC_DL_GreenStrengthIndexCalc := -1.0;  (* 哨兵 -1：组态非法 / Sentinel -1 bad config *)
    RETURN;
END_IF
(* 润滑剂折减因子：含量越高强度越低，下限钳位 0.3 防归零 *)
fLubeFactor := 1.0 - (fLubePct / DL_PCT_BASE) * DL_LUBE_K;
IF fLubeFactor < DL_LF_MIN THEN
    fLubeFactor := DL_LF_MIN;                 (* 下限钳位 [-] / Lower clamp *)
END_IF
(* 压力项非负钳位后开方（开方前判非负） *)
fPressPos := fPressMPa;
IF fPressPos < DL_ZERO THEN
    fPressPos := DL_ZERO;
END_IF
(* 强度指数：sqrt(p) × 增益 × 润滑剂因子 × 密度比，参考密度已过域闸 *)
fStrengthIdx := SQRT(fPressPos) * DL_GAIN * fLubeFactor * (fGreenDens / fDensRef);
(* 脱模安全判定：指数达阈值即可安全脱模 *)
xEjectSafe := fStrengthIdx >= fSafeIdx;
xValid := TRUE;                               (* 链路有效 / Chain valid *)
FC_DL_GreenStrengthIndexCalc := fStrengthIdx; (* 返回强度指数 [-] / Return strength index *)
END_FUNCTION

(* ---- FC_DL_HexChromeTriRatioCalc.st ---- *)
(*
  DL Factory R83 | FC_DL_HexChromeTriRatioCalc
  功能：算六价铬与三价铬浓度比，判定镀液老化并给出需氧化的三价铬过量值。
  开源溯源：无（clean-room 自研，依据公开工艺公式，来源=行业通用公式，许可证=MIT，借鉴点=公式结构）
  规则：R1-R21 全遵守
*)
FUNCTION FC_DL_HexChromeTriRatioCalc : REAL
VAR_INPUT
    fCr6Gpl   : REAL; // 六价铬浓度 [g/L] / Hexavalent chromium concentration [g/L]
    fCr3Gpl   : REAL; // 三价铬浓度 [g/L] / Trivalent chromium concentration [g/L]
    fRatioMin : REAL; // 允许最低六/三比值 [-]/ Minimum allowed hex-to-tri ratio [-]
    fTempC    : REAL; // 槽液温度 [°C] / Bath temperature [degC]
END_VAR
VAR_OUTPUT
    fRatio     : REAL; // 六价/三价比值 [-]/ Hex-to-tri concentration ratio [-]
    fCr3Excess : REAL; // 三价铬过量（需氧化去除量，负值按零）[g/L] / Excess trivalent [g/L]
    xAged      : BOOL; // 老化判定（TRUE=三价累积超限）/ Ageing flag, TRUE = build-up
    xValid     : BOOL; // 计算有效性标志 / Calculation validity flag
END_VAR
VAR
    fCr3Limit : REAL; // 三价铬允许上限 [g/L] / Allowed trivalent ceiling [g/L]
END_VAR
// 出口预置：四出口统一预置，老化标志预置 FALSE（安全侧）
fRatio := 0.0; fCr3Excess := 0.0; xAged := FALSE; xValid := FALSE;
// 非有限拦截 + 量纲自检（R20/R21）
IF NOT (fCr6Gpl > -1.0E30 AND fCr6Gpl < 1.0E30) OR NOT (fCr3Gpl > -1.0E30 AND fCr3Gpl < 1.0E30) OR NOT (fRatioMin > -1.0E30 AND fRatioMin < 1.0E30) OR NOT (fTempC > -1.0E30 AND fTempC < 1.0E30) OR fCr6Gpl <= 0.0 OR fCr3Gpl <= 0.0 OR fRatioMin <= 0.0 THEN
    FC_DL_HexChromeTriRatioCalc := -1.0; RETURN;  // 哨兵 -1：非有限或量纲越界 / Sentinel -1
END_IF
// 比值：六价 ÷ 三价，两者同量纲 g/L 故比值为无量纲；三价分母显式零闸（R4/R21）
IF ABS(fCr3Gpl) > 1.0E-9 THEN       // 三价分母显式零闸 / Explicit zero gate on trivalent
    fRatio := fCr6Gpl / fCr3Gpl;    // 六/三比值 [-]/ Hex-to-tri ratio
ELSE
    fRatio := 0.0;                  // 除零防御缺省 / Divide-by-zero default
END_IF
// 三价上限：由比值下限反算 Cr3 <= Cr6 ÷ 比值下限（g/L ÷ 无量纲 = g/L）
IF ABS(fRatioMin) > 1.0E-9 THEN     // 比值下限分母显式零闸 / Zero gate on ratio lower bound
    fCr3Limit := fCr6Gpl / fRatioMin;   // 三价允许上限 [g/L] / Allowed trivalent ceiling
ELSE
    fCr3Limit := fCr3Gpl;           // 下限非正时按当前值兜底，不产生过量 / Fallback, no excess
END_IF
// 过量：三价实测减允许上限，负值按零（单向语义，不做浓缩回算）
IF fCr3Gpl > fCr3Limit THEN
    fCr3Excess := fCr3Gpl - fCr3Limit;  // 超量部分 [g/L] / Excessive part [g/L]
    xAged      := TRUE;             // 三价累积超限判老化 / Build-up flags ageing
ELSE
    fCr3Excess := 0.0;              // 未超限，过量按零 / Not exceeded, zero
    xAged      := FALSE;            // 比值正常 / Ratio within limit
END_IF
xValid := TRUE; FC_DL_HexChromeTriRatioCalc := fRatio;  // 返回六/三比值 [-] / Return ratio
END_FUNCTION

(* ---- FC_DL_IdleRunRatioCalc.st ---- *)
(*
  ============================================================
  组件名 : FC_DL_IdleRunRatioCalc
  分类   : DL_Process
  功能   : 空转率与浪费电量计算，由总运行时间与加载时间求空转占比及折算电耗
  复杂度 : C1
  版本   : 1.0.0
  作者   : 道莅工业代码库工厂 / R81
  日期   : 2026-11-24
  开源溯源 : clean-room（no upstream）—— 依据公开工程公式自研，未复制任何上游实现
  红线自检 : R1 无GVL/R2 无物理地址/R3 纯IEC/R4 防除零/R5 双语注释
  接口说明 :
      空转时间 = 总运行时间 - 加载时间；空转率 = 空转时间 / 总运行时间 * 100。
      浪费电量 = 空转功率 * 空转时间 / 3600，单位 kWh。
      加载时间超过总运行时间属数据矛盾，本组件判无效，不做负数截断掩盖问题。
  ============================================================
*)
FUNCTION FC_DL_IdleRunRatioCalc : BOOL
VAR_INPUT
    bEnable     : BOOL; // 使能：TRUE 时计算 / Enable: TRUE to compute
    bErr        : BOOL; // 外部故障：TRUE 时立即退出并置结果无效 / External fault: TRUE aborts with invalid result
    rRunTime_s  : REAL; // 总运行时间 [s] / total running time [second]
    rLoadTime_s : REAL; // 加载运行时间 [s] / loaded running time [second]
    rIdleKw     : REAL; // 空转状态功率 [kW] / idle state power [kilowatt]
END_VAR
VAR_OUTPUT
    rIdleTime_s : REAL; // 空转时间 [s] / idle time [second]
    rIdlePct    : REAL; // 空转率，限幅 0~100 [%] / idle ratio clamped to 0 to 100 [percent]
    rWastedKwh  : REAL; // 空转浪费电量 [kWh] / energy wasted while idling [kilowatt hour]
    bValid      : BOOL; // 输出有效：TRUE 表示结果可用 / Output valid
END_VAR
VAR CONSTANT
    DL_R_MAX   : REAL := 3.0E38;  // 实数上界，用于拦截 Inf [无量纲] / real upper bound used to reject infinity [dimensionless]
    DL_EPS     : REAL := 1.0E-12; // 除零判定阈值 [无量纲] / division guard threshold [dimensionless]
    DL_PCT     : REAL := 100.0;   // 百分数换算系数 [无量纲] / percentage scaling factor [dimensionless]
    DL_ZERO    : REAL := 0.0;     // 零值常量 [无量纲] / zero constant [dimensionless]
    DL_S_PER_H : REAL := 3600.0;  // 每小时秒数 [s/h] / seconds per hour [second per hour]
    DL_TOL_S   : REAL := 0.001;   // 时间比较容差 [s] / tolerance of the time comparison [second]
END_VAR
VAR
    _bFin : BOOL := FALSE; // 输入有限性判定结果 / input finiteness verdict
END_VAR

    // 段 1｜出口预置
    rIdleTime_s := 0.0;
    rIdlePct := 0.0;
    rWastedKwh := 0.0;
    bValid := FALSE;
    // 段 2｜使能闸与外部故障闸
    IF NOT bEnable THEN
        RETURN;
    END_IF;
    IF bErr THEN
        RETURN;
    END_IF;
    // 段 3｜非有限闸
    _bFin := (rRunTime_s = rRunTime_s) AND (ABS(rRunTime_s) <= DL_R_MAX) AND (rLoadTime_s = rLoadTime_s) AND (ABS(rLoadTime_s) <= DL_R_MAX) AND (rIdleKw = rIdleKw) AND (ABS(rIdleKw) <= DL_R_MAX);
    IF NOT _bFin THEN
        RETURN;
    END_IF;
    // 段 4｜域闸：总运行时间严格为正，加载时间与空转功率不得为负
    IF (ABS(rRunTime_s) <= DL_EPS) OR (rRunTime_s < DL_ZERO) THEN
        RETURN;
    END_IF;
    IF (rLoadTime_s < DL_ZERO) OR (rIdleKw < DL_ZERO) THEN
        RETURN;
    END_IF;
    // 段 5｜加载时间不得越过总运行时间
    IF rLoadTime_s > (rRunTime_s + DL_TOL_S) THEN
        RETURN;
    END_IF;
    // 段 6｜空转时间
    rIdleTime_s := rRunTime_s - rLoadTime_s;
    IF rIdleTime_s < DL_ZERO THEN
        rIdleTime_s := DL_ZERO;
    END_IF;
    // 段 7｜空转率与浪费电量
    rIdlePct := rIdleTime_s / rRunTime_s * DL_PCT;
    IF rIdlePct < DL_ZERO THEN
        rIdlePct := DL_ZERO;
    END_IF;
    IF rIdlePct > DL_PCT THEN
        rIdlePct := DL_PCT;
    END_IF;
    rWastedKwh := rIdleKw * rIdleTime_s / DL_S_PER_H;
    bValid := TRUE;
    FC_DL_IdleRunRatioCalc := bValid;
END_FUNCTION

(* ---- FC_DL_ImpulseSealDwellCalc.st ---- *)
(*
  DL Factory R83 | FC_DL_ImpulseSealDwellCalc
  功能：按热封面积、膜厚与温升用能量平衡算通电时间，并给出保压冷却时间。
  开源溯源：无（clean-room 自研，依据公开工艺公式，来源=行业通用公式，许可证=MIT，借鉴点=公式结构）
  规则：R1-R21 全遵守
*)
FUNCTION FC_DL_ImpulseSealDwellCalc : REAL
VAR_INPUT
    fSealAreaMm2  : REAL; // 热封有效面积 [mm²] / Effective seal area [mm^2]
    fFilmThickUm  : REAL; // 封合膜总厚度 [µm] / Total film thickness [um]
    fSealTempC    : REAL; // 热封目标温度 [°C] / Seal target temperature [degC]
    fAmbTempC     : REAL; // 环境（初始）温度 [°C] / Ambient initial temperature [degC]
    fHeaterPowerW : REAL; // 热封头有效功率 [W] / Effective sealer power [W]
END_VAR
VAR_OUTPUT
    fHeatTimeMs  : REAL; // 通电加热时间 [ms] / Power-on heating time [ms]
    fDwellTimeMs : REAL; // 保压冷却时间 [ms] / Dwell cooling time [ms]
    xValid       : BOOL; // 计算有效性标志 / Calculation validity flag
END_VAR
VAR
    fMassG    : REAL; // 封合区膜料质量 [g] / Film mass in seal zone [g]
    fEnergyJ  : REAL; // 所需热量 [J] / Required heat energy [J]
    cDensity  : REAL := 0.92; // 膜密度常量 [g/cm³]，已引用（R19）/ Film density [g/cm^3]
    cSpecHeat : REAL := 1.70; // 比热容常量 [J/(g·K)]，已引用（R19）/ Specific heat [J/(g.K)]
    cEff      : REAL := 0.35; // 热效率常量 [-]，已引用（R19）/ Thermal efficiency [-]
END_VAR
// 出口预置：三出口统一预置（R256）
fHeatTimeMs := 0.0; fDwellTimeMs := 0.0; xValid := FALSE;
// 非有限拦截 + 量纲自检 + 温升方向检查（R20/R21）
IF NOT (fSealAreaMm2 > -1.0E30 AND fSealAreaMm2 < 1.0E30) OR NOT (fFilmThickUm > -1.0E30 AND fFilmThickUm < 1.0E30) OR NOT (fSealTempC > -1.0E30 AND fSealTempC < 1.0E30) OR NOT (fAmbTempC > -1.0E30 AND fAmbTempC < 1.0E30) OR NOT (fHeaterPowerW > -1.0E30 AND fHeaterPowerW < 1.0E30) OR fSealAreaMm2 <= 0.0 OR fFilmThickUm <= 0.0 OR fHeaterPowerW <= 0.0 OR fSealTempC <= fAmbTempC THEN
    FC_DL_ImpulseSealDwellCalc := -1.0; RETURN;   // 哨兵 -1：非有限或量纲/温升越界 / Sentinel -1
END_IF
// 质量：mm² × µm × 1E-6 = cm³，再乘 g/cm³ 得 g（量纲自洽：1 µm = 1E-3 mm，故 1E-3 mm³ = 1E-6 cm³）
fMassG := fSealAreaMm2 * fFilmThickUm * 1.0E-6 * cDensity;   // 封合区质量 [g] / Film mass [g]
// 热量：Q = m × c × ΔT，ΔT 为设定与环境之差（K 与 °C 同尺度，故可直接相减）
fEnergyJ := fMassG * cSpecHeat * (fSealTempC - fAmbTempC);   // 所需热量 [J] / Required energy [J]
// 通电时间：J ÷ W = s，×1000 = ms，再除以热效率放大（含热损，故非恒等式）
fHeatTimeMs := (fEnergyJ / fHeaterPowerW) * 1000.0 / cEff;   // 通电时间 [ms] / Heating time [ms]
// 保压时间：取通电时间 40% 加厚膜附加项，保证熔接层冷却定型
fDwellTimeMs := fHeatTimeMs * 0.40 + 50.0 + fFilmThickUm * 0.5; // 保压时间 [ms] / Dwell time [ms]
xValid := TRUE;                                                // 链路有效 / Chain valid
FC_DL_ImpulseSealDwellCalc := fHeatTimeMs;                     // 返回通电时间 [ms] / Return heating time
END_FUNCTION

(* ---- FC_DL_InkViscosityTempComp.st ---- *)
(*
  DL Factory R83 | FC_DL_InkViscosityTempComp
  功能：按温度线性修正系数把实测油墨黏度折算到参考温度，并给出兑稀补偿系数。
  开源溯源：无（clean-room 自研，依据公开工艺公式，来源=行业通用公式，许可证=MIT，借鉴点=公式结构）
  规则：R1-R21 全遵守
*)
FUNCTION FC_DL_InkViscosityTempComp : REAL
VAR_INPUT
    fViscMeas   : REAL; // 实测黏度 [mPa·s] / Measured viscosity [mPa.s]
    fTempMeas   : REAL; // 实测油墨温度 [°C] / Measured ink temperature [degC]
    fTempRef    : REAL; // 参考温度（工艺基准）[°C] / Reference temperature [degC]
    fTempCoeff  : REAL; // 温度系数（每 °C 黏度变化率）[%/°C] / Temperature coefficient [%/degC]
    fViscTarget : REAL; // 目标黏度（工艺设定）[mPa·s] / Target viscosity [mPa.s]
END_VAR
VAR_OUTPUT
    fViscRef    : REAL; // 参考温度下黏度 [mPa·s] / Viscosity at reference temperature [mPa.s]
    fCompFactor : REAL; // 兑稀补偿系数，小于 1 需加溶剂 [-]/ Thinning factor, below 1 means add solvent
    xValid      : BOOL; // 输入有效性（FALSE 时输出为故障缺省）/ Input validity flag
END_VAR
VAR
    fScale : REAL; // 温度修正比例因子 [-] / Temperature correction scale factor
END_VAR
// 出口预置：三出口统一预置，故障拍不残留上拍值（R187/R256）
fViscRef := 0.0; fCompFactor := 0.0; xValid := FALSE;
// 非有限拦截 + 量纲自检：NaN/Inf 与域越界同走故障分支（R20/R21）
IF NOT (fViscMeas > -1.0E30 AND fViscMeas < 1.0E30) OR NOT (fTempMeas > -1.0E30 AND fTempMeas < 1.0E30) OR NOT (fTempRef > -1.0E30 AND fTempRef < 1.0E30) OR NOT (fTempCoeff > -1.0E30 AND fTempCoeff < 1.0E30) OR NOT (fViscTarget > -1.0E30 AND fViscTarget < 1.0E30) OR fViscMeas <= 0.0 OR fTempRef <= -50.0 OR fTempRef > 200.0 THEN
    FC_DL_InkViscosityTempComp := -1.0; RETURN;   // 哨兵 -1：非有限或量纲越界 / Sentinel -1
END_IF
// 温度折算：η(Tref) = η(T) × (1 + k × (Tref - T))，线性工艺近似
fScale := 1.0 + (fTempCoeff / 100.0) * (fTempRef - fTempMeas); // 比例因子 [-] / Scale factor
IF fScale > 0.05 THEN                    // 比例因子下限闸，防负值或近零
    fViscRef := fViscMeas * fScale;      // 参考温度黏度 [mPa·s] / Viscosity at ref temp
ELSE
    fViscRef := fViscMeas;               // 极端温差回退实测值 / Fallback to measured
END_IF
// 补偿系数：目标黏度 ÷ 折算实值，含目标工艺量故非恒等式
IF ABS(fViscRef) > 1.0E-9 THEN           // 分母显式零闸（R4/R21）/ Explicit zero gate
    fCompFactor := fViscTarget / fViscRef;  // 兑稀补偿系数 [-]/ Thinning factor
    xValid      := TRUE;                 // 计算链路有效 / Chain valid
ELSE
    fCompFactor := 0.0;                  // 除零防御缺省 / Divide-by-zero default
END_IF
FC_DL_InkViscosityTempComp := fCompFactor; // 返回兑稀补偿系数 [-]/ Return thinning factor
END_FUNCTION

(* ---- FC_DL_JacketAreaCalc.st ---- *)
(*
  DL Factory R84 | FC_DL_JacketAreaCalc
  功能：由所需换热量与总传热系数算夹套/盘管传热面积，含 LMTD 计算与面积校核
  开源溯源：无（clean-room 自研，依据公开工艺公式，来源=行业通用公式，许可证=MIT，借鉴点=公式结构）
  规则：R1-R16 全遵守
*)
FUNCTION FC_DL_JacketAreaCalc : REAL
VAR_INPUT
    fQDutyKw : REAL := 120.0; // 所需换热量 [kW] / required heat duty [kW]
    fKWm2K : REAL := 350.0; // 总传热系数 [W/(m²·K)] / overall heat transfer coefficient [W/(m^2*K)]
    fThInC : REAL := 90.0; // 热侧进口温度 [℃] / hot side inlet temperature [C]
    fThOutC : REAL := 70.0; // 热侧出口温度 [℃] / hot side outlet temperature [C]
    fTcInC : REAL := 25.0; // 冷侧进口温度 [℃] / cold side inlet temperature [C]
    fTcOutC : REAL := 40.0; // 冷侧出口温度 [℃] / cold side outlet temperature [C]
    fAreaAvailM2 : REAL := 6.0; // 现有可用传热面积（校核用） [m²] / available heat transfer area [m^2]
END_VAR
VAR_OUTPUT
    fLmtd : REAL; // 对数平均温差 [K] / log mean temperature difference [K]
    fQreqKw : REAL; // 所需换热量回显（链路校验） [kW] / required duty echo [kW]
    xValid : BOOL; // 计算结果有效标志 [-] / calculation valid flag [-]
END_VAR
VAR
    fDt1K : REAL; // 端差 1（热进 − 冷出） [K] / terminal difference one [K]
    fDt2K : REAL; // 端差 2（热出 − 冷进） [K] / terminal difference two [K]
    fAreaM2 : REAL; // 所需传热面积 [m²] / required area [m^2]
    xAreaOk : BOOL; // 面积是否满足（A 需求 ≤ 可用） [-] / area adequacy verdict [-]
END_VAR

// 段 1｜出口预置（R256）
FC_DL_JacketAreaCalc := -1.0; // 哨兵返回 -1（无效） [-] / sentinel return -1, invalid [-]
fLmtd := 0.0; // LMTD 预置零 [K] / LMTD preset zero [K]
fQreqKw := 0.0; // 热量回显预置零 [kW] / duty echo preset zero [kW]
xValid := FALSE; // 计算完成前不认结果 [-] / unusable before calculation [-]

// 段 2｜非有限拦截 + 域闸（R4/R20）
IF NOT (fQDutyKw > -1.0E30 AND fQDutyKw < 1.0E30) OR NOT (fKWm2K > -1.0E30 AND fKWm2K < 1.0E30) OR NOT (fThInC > -1.0E30 AND fThInC < 1.0E30) OR NOT (fThOutC > -1.0E30 AND fThOutC < 1.0E30) THEN
    RETURN; // 热量/系数/热侧温度任一非有限即拒算 [-] / any non finite duty, coefficient or hot side rejected [-]
END_IF
IF NOT (fTcInC > -1.0E30 AND fTcInC < 1.0E30) OR NOT (fTcOutC > -1.0E30 AND fTcOutC < 1.0E30) OR NOT (fAreaAvailM2 > -1.0E30 AND fAreaAvailM2 < 1.0E30) THEN
    RETURN; // 冷侧温度或可用面积非有限即拒算 [-] / any non finite cold side or area rejected [-]
END_IF
IF fKWm2K < 1.0E-9 OR fQDutyKw < 0.0 OR fAreaAvailM2 < 0.0 THEN
    RETURN; // K 值正域分母闸 + 热量/面积非负闸 [W/(m²·K), kW, m²] / positive K denominator gate [-]
END_IF

// 段 3｜端差与 LMTD
fDt1K := fThInC - fTcOutC; // ℃ − ℃ = K（温差） / [C] minus [C] = [K]
fDt2K := fThOutC - fTcInC; // ℃ − ℃ = K（温差） / [C] minus [C] = [K]
IF (fDt1K < 1.0E-9) OR (fDt2K < 1.0E-9) THEN
    RETURN; // 任一端差非正：温度交叉或逆流不可行，拒算 [-] / non positive terminal difference rejected [-]
END_IF
IF ABS(fDt1K - fDt2K) < 1.0E-9 THEN
    fLmtd := fDt1K; // 两端差相等时 LMTD 退化为该端差 [K] / degenerate case, LMTD equals the difference [K]
ELSE
    fLmtd := (fDt1K - fDt2K) / LN(fDt1K / fDt2K); // K ÷ 无量纲 = K（K/K 取对数无量纲） / [K] / [-] = [K]
END_IF
IF NOT (fLmtd > 1.0E-9) OR NOT (fLmtd < 1.0E30) THEN
    RETURN; // LMTD 分母闸：必须为正有限值 [K] / LMTD must be positive and finite [K]
END_IF

// 段 4｜面积 A = Q / (K × LMTD)，并与可用面积校核
fAreaM2 := (fQDutyKw * 1000.0) / (fKWm2K * fLmtd); // (kW×1000 = W) ÷ (W/(m²·K)×K) = m² / [kW]×1000 / ([W/(m^2*K)]×[K]) = [m^2]
IF NOT (fAreaM2 > -1.0E30 AND fAreaM2 < 1.0E30) THEN
    RETURN; // 结果非有限再拦一次 [-] / second finiteness gate [-]
END_IF
xAreaOk := fAreaM2 <= fAreaAvailM2; // m² 直比，禁浮点等值 [-] / direct compare of the areas [m^2]
fQreqKw := fQDutyKw; // 回显所需换热量 [kW] / echo the required duty [kW]
xValid := xAreaOk; // 面积不足即判无效（需加大设备或提 K 值） [-] / area shortage voids the result [-]
FC_DL_JacketAreaCalc := fAreaM2; // 返回所需面积 [m²] / return the required area [m^2]
END_FUNCTION

(* ---- FC_DL_JiggerLiquorRatioCalc.st ---- *)
(*
  Name: FC_DL_JiggerLiquorRatioCalc
  Category: DL_Process
  Version: 1.0.0
  Round: R91 / 2026-11-25
  开源溯源：clean-room 自研（族 间歇式溢流染色与丝光整理，ST 开源生态实测 0 命中，无外部代码引入）
  说明：本件与在册 FC_DL_DyeLiquorRatioCalc（由「重量 × 浴比」正算总液量）方向相反，
        本件由「实测液量 ÷ 实测布重」反算实际浴比并做工艺区间判定，输入输出契约无交集，
        属同族内的对偶量而非重复实现（R13 语义查重结论：非重复）。
  功能：1) 实际浴比按「染液体积 / 被染物质量」计算：ratio = V / m，单位 L/kg，
           分母取被染物质量、分子取染液体积，方向固定不可交换（浴比是「每公斤布配多少升液」）。
        2) 工艺区间判定：fRatioLoLkg <= ratio <= fRatioHiLkg 输出 xInBand；
           低于下限判 xRatioLow（浴比过小、布在缸内易打结起皱、染色不匀）；
           高于上限判 xRatioHigh（浴比过大、助剂浪费、污水负荷高）。
        3) 输出偏差量 fDevLkg = ratio − 区间中值，作为补液/排液的前馈修正量
           （正偏差需排液，负偏差需补液，方向由符号给出）。
  边界条件：1) 非有限值闸：四路实值入参先过 NOT(x > -DL_BIG AND x < DL_BIG)，同时拦 NaN 与 Inf，
           命中即闸断实值通路（浴比与偏差强制 0.0），不得只置标志（R19）。
        2) 重量零闸：被染物质量 fFabricKg 必须 > DL_EPS（浴比式的分母）；
           为零时浴比发散，判无效并清零，绝不输出「无穷大浴比」。
        3) 液量非负闸：染液体积不得为负（负体积属液位计反向或组态错），判无效。
        4) 区间域闸：须满足 0.0 < fRatioLoLkg < fRatioHiLkg <= DL_RATIO_HI_LKG，
           否则两级判据重叠或倒置，越域判无效并把偏低位置真（保守侧）。
        5) 判据取原始值（R24）：区间判定使用钳制前的 _fRatioRawLkg，钳制只作用于输出。
        6) 纯函数无状态：补液/排液的累计与联锁由上层染缸批次序 FB 承担。
  量纲自证：ratio = (L)/(kg) = L/kg，与两个区间阈同量纲，可直接比较；
           fDevLkg = (L/kg) − (L/kg) = L/kg，减法两侧同量纲，量纲合法。
  修订历史 Revision :
    2026-11-25  v1.0.0  R91 首版
*)

FUNCTION FC_DL_JiggerLiquorRatioCalc : BOOL
VAR_INPUT
    fLiquorVolL      : REAL;   // 染液实际体积 [L] / Actual dye liquor volume [L]
    fFabricKg        : REAL;   // 被染物（布卷）质量 [kg] / Fabric batch mass [kg]
    fRatioLoLkg      : REAL;   // 工艺浴比下限 [L/kg] / Process liquor ratio low limit [L/kg]
    fRatioHiLkg      : REAL;   // 工艺浴比上限 [L/kg] / Process liquor ratio high limit [L/kg]
END_VAR
VAR_OUTPUT
    fRatioLkg        : REAL;   // 实际浴比 [L/kg] / Actual liquor ratio [L/kg]
    fDevLkg          : REAL;   // 相对区间中值的偏差 [L/kg] / Deviation from the band mid value [L/kg]
    xRatioLow        : BOOL;   // 低于下限标志 [bool] / Below the low limit flag [bool]
    xRatioHigh       : BOOL;   // 高于上限标志 [bool] / Above the high limit flag [bool]
    xValid           : BOOL;   // 计算有效标志 [bool] / Calculation valid flag [bool]
END_VAR
VAR
    _fRatioRawLkg    : REAL;   // 钳制前的原始浴比 [L/kg] / Raw liquor ratio before limiting [L/kg]
    _fMidLkg         : REAL;   // 区间中值 [L/kg] / Mid value of the band [L/kg]
    _fDevRawLkg      : REAL;   // 钳制前的原始偏差 [L/kg] / Raw deviation before limiting [L/kg]
END_VAR
VAR CONSTANT
    DL_EPS           : REAL := 1.0E-9;    // 数值零闸阈值 [-] / Numeric zero gate threshold [-]
    DL_BIG           : REAL := 1.0E12;    // 非有限值闸量级上限 [-] / Finiteness gate magnitude [-]
    DL_HALF          : REAL := 0.5;       // 区间中值折算系数 [-] / Band mid-point factor [-]
    DL_RATIO_HI_LKG  : REAL := 100.0;     // 浴比物理上限 [L/kg] / Liquor ratio physical upper bound [L/kg]
    DL_DEV_SPAN      : REAL := 100.0;     // 偏差钳制跨度 [L/kg] / Deviation clamp span [L/kg]
END_VAR

(* —— 段 1：非有限值闸（R19：闸断实值通路） —— *)
IF NOT (fLiquorVolL > -DL_BIG AND fLiquorVolL < DL_BIG)
   OR NOT (fFabricKg > -DL_BIG AND fFabricKg < DL_BIG)
   OR NOT (fRatioLoLkg > -DL_BIG AND fRatioLoLkg < DL_BIG)
   OR NOT (fRatioHiLkg > -DL_BIG AND fRatioHiLkg < DL_BIG) THEN
    fRatioLkg := 0.0;                       // 输出强制 0.0，切断污染源 / Force zero, cut polluted path
    fDevLkg := 0.0;                         // 偏差强制 0.0 / Deviation forced to zero
    xRatioLow := TRUE;                      // 失效侧按偏低处理（保守侧：提示补液）
    xRatioHigh := FALSE;                    // 失效侧偏高位保持假 / High flag stays false
    xValid := FALSE;                        // 有效位清零 / Validity cleared
    FC_DL_JiggerLiquorRatioCalc := FALSE;   // 返回码与有效位同源 / Return mirrors validity
    RETURN;                                 // 立即退出 / Immediate exit
END_IF

(* —— 段 2：重量零闸与区间域闸（分母为布重） —— *)
IF (fFabricKg <= DL_EPS)                                          // 布重不可为零
   OR (fLiquorVolL < 0.0)                                         // 液量不得为负
   OR (fRatioLoLkg <= 0.0)                                        // 区间下限必须为正
   OR (fRatioHiLkg <= fRatioLoLkg)                                // 区间必须有效（hi > lo）
   OR (fRatioHiLkg > DL_RATIO_HI_LKG) THEN                        // 上限须在物理域内
    fRatioLkg := 0.0;                       // 布重为零即不可算 / No mass, no ratio
    fDevLkg := 0.0;                         // 偏差不可算 / Deviation not computable
    xRatioLow := TRUE;                      // 按偏低处理（保守侧）/ Treat as low
    xRatioHigh := FALSE;                    // 偏高位保持假 / High flag stays false
    xValid := FALSE;                        // 判无效 / Invalid
    FC_DL_JiggerLiquorRatioCalc := FALSE;   // 返回码同步 / Return synchronised
    RETURN;                                 // 提前退出 / Early exit
END_IF

(* —— 段 3：主算式（不钳制，先出原始值供段 4 判据使用，R24） —— *)
_fRatioRawLkg := fLiquorVolL / fFabricKg;                                         // 实际浴比 [L/kg]
_fMidLkg := (fRatioLoLkg + fRatioHiLkg) * DL_HALF;                                // 区间中值 [L/kg]
_fDevRawLkg := _fRatioRawLkg - _fMidLkg;                                          // 相对中值偏差 [L/kg]

(* —— 段 4：判据（取原始值；单点 BOOL 聚合避免多处赋 FALSE 覆盖） —— *)
xRatioLow := (_fRatioRawLkg < fRatioLoLkg);                                       // 低于下限
xRatioHigh := (_fRatioRawLkg > fRatioHiLkg);                                      // 高于上限
xValid := (_fRatioRawLkg >= 0.0)                                                  // 浴比不得为负
          AND (_fRatioRawLkg <= DL_RATIO_HI_LKG)                                  // 不超物理上限（量级异常）
          AND (_fMidLkg > 0.0);                                                   // 中值必须为正（区间已验）

(* —— 段 5：输出单点写盘（钳制到物理域内，判定结果已在段 4 定案） —— *)
fRatioLkg := LIMIT(0.0, _fRatioRawLkg, DL_RATIO_HI_LKG);                          // 浴比钳物理域 [L/kg]
fDevLkg := LIMIT(-DL_DEV_SPAN, _fDevRawLkg, DL_DEV_SPAN);                          // 偏差钳物理域 [L/kg]
FC_DL_JiggerLiquorRatioCalc := xValid;                                            // 返回码：TRUE = 计算可信

END_FUNCTION

(* ---- FC_DL_JiggerRampRateCalc.st ---- *)
(*
  Name: FC_DL_JiggerRampRateCalc
  Category: DL_Process
  Version: 1.0.0
  Round: R91 / 2026-11-25
  开源溯源：clean-room 自研（族 间歇式溢流染色与丝光整理，ST 开源生态实测 0 命中，无外部代码引入）
  功能：1) 升温速率按「目标与当前的温差 / 设定升温时间」计算：rate = dT / t，单位 degC/min，
           分母为设定升温时长（分钟），故无需再乘 60，避免二次折算引入量纲错误。
        2) 纤维允许速率上限校验：rate > fRateMaxKmin 输出 xRateOver（超纤维允许速率），
           这是「快速升温导致染料上染过快、产生色花与折痕」的直接判据；
           对涤纶等疏水纤维该上限通常只有 1.0 ~ 1.5 degC/min。
        3) 输出温差 fDeltaK 与速率 fRateKmin 两个量：温差供设备能力校核
           （蒸汽阀全开能否在设定时间内完成），速率供工艺合规校核。
  边界条件：1) 非有限值闸：四路实值入参先过 NOT(x > -DL_BIG AND x < DL_BIG)，同时拦 NaN 与 Inf，
           命中即闸断实值通路（速率与温差强制 0.0 且置超限位，保守侧），不得只置标志（R19）。
        2) 时间零闸：设定升温时间 fRampMin 必须 > DL_EPS（速率式的分母），
           为零时速率发散，判无效并清零，绝不输出「无穷快升温」。
        3) 温差方向闸：目标温度必须高于当前温度（dT > 0）；dT <= 0 说明这不是升温段
           （可能是降温或保温），本件不适用，判无效而不输出负速率。
        4) 上限域闸：fRateMaxKmin 必须落在 (0.0, DL_RATE_ABS_HI] 内，越域判无效（上限未组态则判据恒假）。
        5) 判据取原始值（R24）：超上限判定使用钳制前的 _fRateRawKmin，钳制只作用于输出。
        6) 纯函数无状态：实际速率（由温度微分测得）与设定速率的比对由上层温控 FB 承担。
  量纲自证：rate = (degC)/(min) = degC/min（温差尺度上与 K/min 等价），
           与 fRateMaxKmin 同量纲，可直接比较；fDeltaK = (degC) − (degC) = K。
  修订历史 Revision :
    2026-11-25  v1.0.0  R91 首版
*)

FUNCTION FC_DL_JiggerRampRateCalc : BOOL
VAR_INPUT
    fStartC          : REAL;   // 当前（起点）染液温度 [degC] / Current dye liquor temperature [degC]
    fTargetC         : REAL;   // 目标染液温度 [degC] / Target dye liquor temperature [degC]
    fRampMin         : REAL;   // 设定升温时长 [min] / Planned heating duration [min]
    fRateMaxKmin     : REAL;   // 纤维允许升温速率上限 [K/min] / Fibre-permitted heating rate limit [K/min]
END_VAR
VAR_OUTPUT
    fRateKmin        : REAL;   // 设定升温速率 [K/min] / Planned heating rate [K/min]
    fDeltaK          : REAL;   // 需升高的温差 [K] / Temperature difference to be raised [K]
    xRateOver        : BOOL;   // 超纤维允许速率标志 [bool] / Over fibre-permitted rate flag [bool]
    xValid           : BOOL;   // 计算有效标志 [bool] / Calculation valid flag [bool]
END_VAR
VAR
    _fDeltaRawK      : REAL;   // 未钳制的温差 [K] / Unclamped temperature difference [K]
    _fRateRawKmin    : REAL;   // 钳制前的原始速率 [K/min] / Raw rate before limiting [K/min]
END_VAR
VAR CONSTANT
    DL_EPS           : REAL := 1.0E-9;    // 数值零闸阈值 [-] / Numeric zero gate threshold [-]
    DL_BIG           : REAL := 1.0E12;    // 非有限值闸量级上限 [-] / Finiteness gate magnitude [-]
    DL_RATE_ABS_HI   : REAL := 50.0;      // 升温速率绝对物理上限 [K/min] / Absolute rate upper bound [K/min]
    DL_T_SPAN        : REAL := 500.0;     // 温度量级闸跨度 [degC] / Temperature magnitude gate span [degC]
END_VAR

(* —— 段 1：非有限值闸（R19：闸断实值通路；失效侧置超限位，保守侧） —— *)
IF NOT (fStartC > -DL_BIG AND fStartC < DL_BIG)
   OR NOT (fTargetC > -DL_BIG AND fTargetC < DL_BIG)
   OR NOT (fRampMin > -DL_BIG AND fRampMin < DL_BIG)
   OR NOT (fRateMaxKmin > -DL_BIG AND fRateMaxKmin < DL_BIG) THEN
    fRateKmin := 0.0;                       // 输出强制 0.0，切断污染源 / Force zero, cut polluted path
    fDeltaK := 0.0;                         // 温差强制 0.0 / Difference forced to zero
    xRateOver := TRUE;                      // 失效侧按超限处理（保守侧：禁止放行升温）
    xValid := FALSE;                        // 有效位清零 / Validity cleared
    FC_DL_JiggerRampRateCalc := FALSE;      // 返回码与有效位同源 / Return mirrors validity
    RETURN;                                 // 立即退出 / Immediate exit
END_IF

(* —— 段 2：时间零闸与上限域闸（分母为设定升温时长） —— *)
IF (fRampMin <= DL_EPS)                                           // 升温时长不可为零
   OR (fRateMaxKmin <= 0.0)                                       // 上限必须为正
   OR (fRateMaxKmin > DL_RATE_ABS_HI)                             // 上限不得超物理上限
   OR (ABS(fStartC) > DL_T_SPAN)                                  // 起点温度量级闸
   OR (ABS(fTargetC) > DL_T_SPAN) THEN                            // 目标温度量级闸
    fRateKmin := 0.0;                       // 时长为零即不可算 / No duration, no rate
    fDeltaK := 0.0;                         // 温差不可用 / Difference not usable
    xRateOver := TRUE;                      // 按超限处理（保守侧）/ Treat as over the limit
    xValid := FALSE;                        // 判无效 / Invalid
    FC_DL_JiggerRampRateCalc := FALSE;      // 返回码同步 / Return synchronised
    RETURN;                                 // 提前退出 / Early exit
END_IF

(* —— 段 3：主算式（不钳制，先出原始值供段 4 判据使用，R24） —— *)
_fDeltaRawK := fTargetC - fStartC;                                                // 需升温温差 [K]
_fRateRawKmin := _fDeltaRawK / fRampMin;                                          // 设定升温速率 [K/min]

(* —— 段 4：判据（取原始值；单点 BOOL 聚合避免多处赋 FALSE 覆盖） —— *)
xRateOver := (_fRateRawKmin > fRateMaxKmin);                                      // 超纤维允许速率
xValid := (_fDeltaRawK > 0.0)                                                     // 必须是升温段（方向固定）
          AND (_fRateRawKmin >= 0.0)                                              // 速率不得为负
          AND (_fRateRawKmin <= DL_RATE_ABS_HI);                                  // 不超绝对物理上限

(* —— 段 5：输出单点写盘（钳制到物理域内，判定结果已在段 4 定案） —— *)
fRateKmin := LIMIT(0.0, _fRateRawKmin, DL_RATE_ABS_HI);                           // 速率钳物理域 [K/min]
fDeltaK := LIMIT(0.0, _fDeltaRawK, DL_T_SPAN);                                    // 温差钳物理域 [K]
FC_DL_JiggerRampRateCalc := xValid;                                               // 返回码：TRUE = 计算可信

END_FUNCTION

(* ---- FC_DL_KegFillingCounterPressureCalc.st ---- *)
// FC_DL_KegFillingCounterPressureCalc v1.0.0
// 开源溯源：clean-room 自研（族 DL_Process，ST 生态实测 0 命中，无外部代码引入）
(*
  功能: 桶装背压：饱和压 = 亨利常数·CO2 体积倍数·(1 + 0.02·(T − 10))（温度线性修正为工程近似，
        非严格亨利温度指数式）；静压 = ρ·g·h/1e5 [bar]；背压 = 饱和压 + 静压 + 0.2 bar 裕量。
  邻件/码位: 用酒温与 CO2 目标定背压，与 FC_DL_BeerCoolingLoadCalc 的降温工序衔接；
             16#0002_9237 = 非有限、CO2 倍数/亨利常数/密度非正、高度为负或背压超 6 bar。
*)
FUNCTION FC_DL_KegFillingCounterPressureCalc : REAL
VAR_INPUT
    fBeerTemp : REAL := 4.0;        // 酒温 [°C] / Beer temperature [degC]
    fCO2Vol   : REAL := 2.5;        // 目标 CO2 体积倍数 [-]，域 > 0 / CO2 volumes
    fHenryK   : REAL := 0.65;       // 亨利常数 [bar]，域 > 0 / Henry constant [bar]
    fHeight   : REAL := 3.0;        // 液柱高度 [m]，域 >= 0 / Liquid column height [m]
    fDensity  : REAL := 1010.0;     // 啤酒密度 [kg/m³]，域 > 0 / Beer density [kg/m^3]
END_VAR
VAR_OUTPUT
    fCounterPressure : REAL;        // 背压设定 [bar]，工艺界 6.0 / Counter pressure [bar]
    bValid           : BOOL;        // 结果有效回执 [-] / Result validity receipt
    uErrorId         : UDINT;       // 事件码，0 = 无事件 / Event code
END_VAR
VAR
    fSatPress : REAL := 0.0;        // 饱和压 [bar] / Saturation pressure [bar]
    fStatic   : REAL := 0.0;        // 液柱静压 [bar] / Hydrostatic pressure [bar]
END_VAR
// 段 0：全路径出口安全缺省 / Safe defaults on all outlets
fCounterPressure := 0.0;            // 背压缺省零 / Counter pressure default zero
bValid := FALSE;                    // 有效回执预清 / Validity preset clear
uErrorId := 16#0000;                // 事件码预清 / Event code preset clear
FC_DL_KegFillingCounterPressureCalc := 0.0;     // 返回值缺省零（镜像背压）/ Return default zero
// 段 1：非有限闸（五入参全枚举）/ Non-finite gate over all inputs
IF (fBeerTemp <> fBeerTemp) OR (fCO2Vol <> fCO2Vol) OR (fHenryK <> fHenryK)
   OR (fHeight <> fHeight) OR (fDensity <> fDensity)
   OR (ABS(fBeerTemp) >= 3.0E38) OR (ABS(fCO2Vol) >= 3.0E38) OR (ABS(fHenryK) >= 3.0E38)
   OR (ABS(fHeight) >= 3.0E38) OR (ABS(fDensity) >= 3.0E38) THEN
    uErrorId := 16#0002_9237;   // 入参非有限拒收 / Non-finite input reject
    RETURN;
END_IF
// 段 2：域闸（CO2 倍数与亨利常数非正拒收 + 密度正 + 高度非负，R4）/ Domain gate
IF (fCO2Vol <= 1.0E-6) OR (fHenryK <= 1.0E-6) THEN
    uErrorId := 16#0002_9237;   // CO2 倍数或亨利常数非正 / Non-positive CO2 or Henry constant
    RETURN;
END_IF
IF fDensity <= 1.0E-6 THEN
    uErrorId := 16#0002_9237;   // 密度非正，静压不可解 / Non-positive density
    RETURN;
END_IF
IF fHeight < 0.0 THEN
    uErrorId := 16#0002_9237;   // 液柱高度为负 / Negative liquid height
    RETURN;
END_IF
// 段 3：主计算（饱和压 + 静压 + 裕量）/ Main computation
fSatPress := fHenryK * fCO2Vol * (1.0 + 0.02 * (fBeerTemp - 10.0));     // 饱和压 [bar] / Saturation
fStatic := fDensity * 9.81 * fHeight / 1.0E5;                           // 静压 [bar] / Hydrostatic
fCounterPressure := fSatPress + fStatic + 0.2;                          // 背压 [bar] / Counter pressure
// 段 4：出口闸（非有限复核 + 6 bar 工艺界判定）/ Outlet gate
IF (fCounterPressure <> fCounterPressure) OR (ABS(fCounterPressure) >= 3.0E38)
   OR (fCounterPressure <= 0.0) THEN
    fCounterPressure := 0.0;    // 复核失败回缺省 / Fallback on recheck failure
    uErrorId := 16#0002_9237;   // 出口复核拒收 / Output recheck reject
    RETURN;
END_IF
IF fCounterPressure > 6.0 THEN
    uErrorId := 16#0002_9237;   // 信息级：背压超 6 bar（桶耐压风险）/ Info: pressure above bound
    RETURN;                     // bValid 保持 FALSE / Validity stays false
END_IF
bValid := TRUE;                 // 有效回执 / Validity receipt
FC_DL_KegFillingCounterPressureCalc := fCounterPressure;    // 返回值镜像背压 / Return mirrors pressure
END_FUNCTION

(* ---- FC_DL_KilnBypassRatioCalc.st ---- *)
(*
  Name: FC_DL_KilnBypassRatioCalc
  Category: DL_Process
  Version: 1.0.0
  Round: R91 / 2026-11-25
  开源溯源：clean-room 自研（族 水泥窑篦冷机与预热器，ST 开源生态实测 0 命中，无外部代码引入）
  功能：1) 窑尾旁路放风比 = 旁路抽风量 / 窑尾总风量 * 100，分母取窑尾总风量（含旁路），
           方向固定不可交换：分子是被抽走的那一支，分母是全量。
        2) 碱氯负荷约束下的推荐区间由 fRatioLoPct / fRatioHiPct 两个组态引脚给出，
           低于下限意味着碱氯循环富集无法抑制，高于下限则热耗与废气处理负担过大；
           输出 xBelowBand / xAboveBand 两个方向判据，供上层决定增开放风或收小放风。
        3) 偏差量 fDevPct 给出与区间中值的偏移，正值为偏高、负值为偏低，
           作为放风阀 PID 的前馈修正量使用（不做积分，积分在阀门回路内）。
  边界条件：1) 非有限值闸：四路实值入参先过 NOT(x > -DL_BIG AND x < DL_BIG)，同时拦 NaN 与 Inf，
           命中即闸断实值通路（全部输出强制 0.0），不得只置标志（R19）。
        2) 分母零闸：窑尾总风量 |fKilnTailNm3h| <= DL_EPS 时不做除法，判无效并清零全部输出。
        3) 物理域闸：旁路风量与总风量均不得为负；旁路风量不得大于总风量（超出守恒判无效）；
           推荐区间须满足 0.0 <= lo < hi <= 100.0，否则视为组态错误判无效，不钳制。
        4) 判据取原始值（R24）：区间判定使用钳制前的 _fRatioRawPct，不得先钳再判（否则判据恒真）。
        5) 物理域钳制：放风比钳 0.0 ~ 100.0 %；偏差钳 -100.0 ~ +100.0 %。
        6) 纯函数无状态：区间带内的迟滞与放风阀动作延时由下游回路承担，本件不做回差。
  量纲自证：fBypassPct = (Nm3/h)/(Nm3/h)*100 = 无因次百分数 [%]；
           fDevPct = (无因次百分数) − (无因次百分数) = 无因次百分数 [%]，减法两侧同量纲，量纲合法。
  修订历史 Revision :
    2026-11-25  v1.0.0  R91 首版
*)

FUNCTION FC_DL_KilnBypassRatioCalc : BOOL
VAR_INPUT
    fBypassNm3h      : REAL;   // 窑尾旁路放风量 [Nm3/h] / Kiln-tail bypass air flow [Nm3/h]
    fKilnTailNm3h    : REAL;   // 窑尾总风量（含旁路）[Nm3/h] / Total kiln-tail gas flow, bypass included [Nm3/h]
    fRatioLoPct      : REAL;   // 碱氯约束推荐区间下限 [%] / Recommended band low limit, alkali-chloride [%]
    fRatioHiPct      : REAL;   // 碱氯约束推荐区间上限 [%] / Recommended band high limit, alkali-chloride [%]
END_VAR
VAR_OUTPUT
    fBypassPct       : REAL;   // 旁路放风比 [%] / Bypass air ratio [%]
    fDevPct          : REAL;   // 相对区间中值的偏差 [%] / Deviation from the band mid value [%]
    xBelowBand       : BOOL;   // 低于推荐区间标志 [bool] / Below recommended band flag [bool]
    xAboveBand       : BOOL;   // 高于推荐区间标志 [bool] / Above recommended band flag [bool]
    xValid           : BOOL;   // 计算有效标志 [bool] / Calculation valid flag [bool]
END_VAR
VAR
    _fRatioRawPct    : REAL;   // 钳制前的原始放风比 [%] / Raw bypass ratio before limiting [%]
    _fMidPct         : REAL;   // 推荐区间中值 [%] / Mid value of the recommended band [%]
    _fDevRawPct      : REAL;   // 钳制前的原始偏差 [%] / Raw deviation before limiting [%]
END_VAR
VAR CONSTANT
    DL_EPS           : REAL := 1.0E-9;    // 数值零闸阈值 [-] / Numeric zero gate threshold [-]
    DL_BIG           : REAL := 1.0E12;    // 非有限值闸量级上限 [-] / Finiteness gate magnitude [-]
    DL_PCT           : REAL := 100.0;     // 百分比换算因子 [%] / Percent conversion factor [%]
    DL_HALF          : REAL := 0.5;       // 区间中值折算系数 [-] / Band mid-point factor [-]
    DL_DEV_LO_PCT    : REAL := -100.0;    // 偏差物理下限 [%] / Deviation physical low [%]
    DL_DEV_HI_PCT    : REAL := 100.0;     // 偏差物理上限 [%] / Deviation physical high [%]
END_VAR

(* —— 段 1：非有限值闸（R19：闸断实值通路） —— *)
IF NOT (fBypassNm3h > -DL_BIG AND fBypassNm3h < DL_BIG)
   OR NOT (fKilnTailNm3h > -DL_BIG AND fKilnTailNm3h < DL_BIG)
   OR NOT (fRatioLoPct > -DL_BIG AND fRatioLoPct < DL_BIG)
   OR NOT (fRatioHiPct > -DL_BIG AND fRatioHiPct < DL_BIG) THEN
    fBypassPct := 0.0;                      // 输出强制 0.0，切断污染源 / Force zero, cut polluted path
    fDevPct := 0.0;                         // 偏差强制 0.0 / Deviation forced to zero
    xBelowBand := FALSE;                    // 失效侧区间位保持假 / Band flags stay false
    xAboveBand := FALSE;                    // 失效侧区间位保持假 / Band flags stay false
    xValid := FALSE;                        // 有效位清零 / Validity cleared
    FC_DL_KilnBypassRatioCalc := FALSE;     // 返回码与有效位同源 / Return mirrors validity
    RETURN;                                 // 立即退出 / Immediate exit
END_IF

(* —— 段 2：分母零闸（分母为窑尾总风量） —— *)
IF ABS(fKilnTailNm3h) <= DL_EPS THEN
    fBypassPct := 0.0;                      // 无总风量即无放风比 / No total flow, no ratio
    fDevPct := 0.0;                         // 偏差不可算 / Deviation not computable
    xBelowBand := FALSE;                    // 区间位保持假 / Band flags stay false
    xAboveBand := FALSE;                    // 区间位保持假 / Band flags stay false
    xValid := FALSE;                        // 判无效 / Invalid
    FC_DL_KilnBypassRatioCalc := FALSE;     // 返回码同步 / Return synchronised
    RETURN;                                 // 提前退出 / Early exit
END_IF

(* —— 段 3：主算式（不钳制，先出原始值供段 4 判据使用，R24） —— *)
_fRatioRawPct := fBypassNm3h / fKilnTailNm3h * DL_PCT;                            // 原始放风比 [%]
_fMidPct := (fRatioLoPct + fRatioHiPct) * DL_HALF;                                // 区间中值 [%]
_fDevRawPct := _fRatioRawPct - _fMidPct;                                          // 相对中值偏差 [%]

(* —— 段 4：判据（取原始值；单点 BOOL 聚合避免多处赋 FALSE 覆盖） —— *)
xBelowBand := (_fRatioRawPct < fRatioLoPct);                                      // 低于推荐下限
xAboveBand := (_fRatioRawPct > fRatioHiPct);                                      // 高于推荐上限
xValid := (fBypassNm3h >= 0.0)                                                    // 旁路风量不得为负
          AND (fKilnTailNm3h > 0.0)                                               // 总风量必须为正
          AND (fBypassNm3h <= fKilnTailNm3h)                                      // 旁路不得大于总量（守恒）
          AND (fRatioLoPct >= 0.0)                                                // 区间下限不得为负
          AND (fRatioHiPct > fRatioLoPct)                                         // 区间必须有效（hi > lo）
          AND (fRatioHiPct <= DL_PCT)                                             // 区间上限不得超过 100 %
          AND (_fRatioRawPct >= 0.0);                                             // 放风比不得为负

(* —— 段 5：输出单点写盘（钳制到物理域内，判定结果已在段 4 定案） —— *)
fBypassPct := LIMIT(0.0, _fRatioRawPct, DL_PCT);                                   // 放风比钳 0..100 [%]
fDevPct := LIMIT(DL_DEV_LO_PCT, _fDevRawPct, DL_DEV_HI_PCT);                        // 偏差钳 -100..+100 [%]
FC_DL_KilnBypassRatioCalc := xValid;                                               // 返回码：TRUE = 计算可信

END_FUNCTION

(* ---- FC_DL_LamellaAreaCalc.st ---- *)
(*
  道莅工业代码库 / Daoli Industrial ST Library
  组件: FC_DL_LamellaAreaCalc
  分类: DL_Process
  开源溯源: 无（clean-room 工程公式自研；参考公开工艺计算公式，未复制任何受版权保护代码）
  许可证: 本项目自有 (MIT)
  功能: 斜板（斜管）沉淀区投影面积计算，按颗粒沉降速度与板倾角余弦折算并加余量系数
*)
FUNCTION FC_DL_LamellaAreaCalc : BOOL
VAR_INPUT
    rFlowM3h : REAL; // 处理水量 [m3/h] / treated water flow
    rVsMmS : REAL; // 设计颗粒沉降速度 [mm/s] / design particle settling velocity
    rCosTheta : REAL; // 板面与水平面夹角的余弦 [-]，如 60° ≈ 0.5 / cosine of plate inclination
    rAreaSafety : REAL; // 面积余量系数 [-]，典型 1.2~1.5 / area safety factor, typically 1.2~1.5
END_VAR
VAR_OUTPUT
    rAreaM2 : REAL; // 所需斜板投影面积 [m2] / required projected plate area
    bValid : BOOL; // 结果有效位 [-] / result valid flag
    iErrCode : INT; // 事件码 0=正常 1=沉降速度非法 2=倾角过大 3=余量系数非法 4=结果非有限 / event code
END_VAR
VAR CONSTANT
    rSecPerHour : REAL := 3600.0; // 每小时秒数 [s/h] / seconds per hour
    rMmToM : REAL := 0.001; // 毫米转米系数 [m/mm] / millimetre to metre factor
    rCosMin : REAL := 0.1; // 可用余弦下限（倾角过大判据）[-] / minimum usable cosine
    rCosMax : REAL := 1.0; // 余弦物理上限（水平板）[-] / physical ceiling of cosine
END_VAR
VAR
    rFlowM3s : REAL; // 处理水量 [m3/s] / flow in cubic metres per second
    rVsMs : REAL; // 沉降速度 [m/s] / settling velocity in m/s
    rCosUse : REAL; // 生效余弦（上限已钳）[-] / effective cosine, capped at one
    rAreaRaw : REAL; // 未限幅面积 [m2] / unlimited area
END_VAR

    // —— 段 0：全路径预清 —— //
    rFlowM3s := 0.0;
    rVsMs := 0.0;
    rCosUse := 0.0;
    rAreaRaw := 0.0;
    rAreaM2 := 0.0;
    bValid := FALSE;
    iErrCode := 0;
    FC_DL_LamellaAreaCalc := FALSE;
    // —— 段 1：分母闸（沉降速度必须为正） —— //
    IF rVsMmS <= 0.0 THEN
        iErrCode := 1; // 沉降速度非正，面积无定义 / non-positive settling velocity, area undefined
        RETURN;
    END_IF;
    IF rCosTheta <= rCosMin THEN
        iErrCode := 2; // 倾角过大（余弦过小），斜板失效 / inclination too steep, plates ineffective
        RETURN;
    END_IF;
    IF rAreaSafety <= 0.0 THEN
        iErrCode := 3; // 余量系数非法 / invalid safety factor
        RETURN;
    END_IF;
    // —— 段 2：单位归一 [m3/h]->[m3/s]、[mm/s]->[m/s] —— //
    rFlowM3s := rFlowM3h / rSecPerHour; // 水量 [m3/s] / flow in m3/s
    rVsMs := rVsMmS * rMmToM; // 沉速 [m/s] / velocity in m/s
    // —— 段 3：余弦物理上限钳位（cos 不得大于 1） —— //
    IF rCosTheta > rCosMax THEN
        rCosUse := rCosMax; // 超 1 视为水平板 / clamp to horizontal plate
    ELSE
        rCosUse := rCosTheta;
    END_IF;
    // —— 段 4：量纲链 (m3/s)/((m/s)*(-)) = m2 —— //
    rAreaRaw := rFlowM3s / (rVsMs * rCosUse) * rAreaSafety; // 斜板面积 [m2] / lamella area
    IF ABS(rAreaRaw) > 1.0E15 THEN
        iErrCode := 4; // 结果非有限，强制归零 / non-finite result, forced to zero
        RETURN;
    END_IF;
    IF rAreaRaw < 0.0 THEN
        rAreaM2 := 0.0; // 负流量防御 / negative flow guard
    ELSE
        rAreaM2 := rAreaRaw;
    END_IF;
    bValid := TRUE;
    FC_DL_LamellaAreaCalc := TRUE;
END_FUNCTION

(* ---- FC_DL_LeafConditioningMoistureCalc.st ---- *)
(*
 * FC_DL_LeafConditioningMoistureCalc | C2 | DL_Process
 * 功能：松散回潮加水量的计算（干物料守恒，含蒸汽凝结水计入总加水量）       单位：流量 [kg/h]、含水率 [%]
 * 工况边界：入口含水率与出口含水率须在 0~100 %，出口不得达 100 %（入分母）；出口含水率低于入口时判为干燥工况，加水量按 0 发布并置信息位；蒸汽量按全部凝结计入总加水（不区分排汽损失）
 * 代数值回代：G=6000 kg/h、w1=12 %、w2=18 %、蒸汽 0 → Gd=6000×88/100=5280 kg/h；Wadd=5280×6/82=386.3 kg/h；总加水=386.3 kg/h（量纲自洽）
 * 开源溯源：clean-room 自研，未复制任何第三方代码（无外部来源）
 *)
FUNCTION FC_DL_LeafConditioningMoistureCalc : BOOL
VAR_INPUT
    rFeedKgH     : REAL := 6000.0;   // 入口叶片流量（湿基）| inlet leaf mass flow, wet basis [kg/h]
    rMoistInPct  : REAL := 12.0;     // 入口含水率 | inlet moisture [%]
    rMoistOutPct : REAL := 18.0;     // 出口含水率目标 | outlet moisture target [%]
    rSteamKgH    : REAL;             // 直接蒸汽流量（全部凝结计入）| direct steam flow, fully condensed [kg/h]
END_VAR
VAR_OUTPUT
    rWaterAddKgH   : REAL;           // 达到出口水分所需加水量 | water needed to reach the outlet moisture [kg/h]
    rTotalWaterKgH : REAL;           // 总加水量（含蒸汽凝结水）| total water including the condensed steam [kg/h]
    rDryMatterKgH  : REAL;           // 绝干物料流量 | dry matter mass flow [kg/h]
    xReverseMoist  : BOOL;           // 出口水分低于入口（干燥工况，信息级）| outlet below inlet, informational
    xValid         : BOOL;           // 输出有效 | outputs valid
END_VAR
VAR
    xFinG    : BOOL;                 // 入口流量有限性 | inlet flow is finite
    xFinW1   : BOOL;                 // 入口水分有限性 | inlet moisture is finite
    xFinW2   : BOOL;                 // 出口水分有限性 | outlet moisture is finite
    xFinStm  : BOOL;                 // 蒸汽流量有限性 | steam flow is finite
    rDenPct  : REAL;                 // 分母 (100−w2) | denominator 100 minus w2 [%]
END_VAR
VAR CONSTANT
    DL_LCM_PCT_MAX : REAL := 100.0;  // 含水率上限 | upper moisture limit [%]
    DL_LCM_DEN_MIN : REAL := 1.0E-6; // 除零保护阈值 | division guard threshold [%]
END_VAR

// 段1｜非有限闸（R19）
xFinG := (rFeedKgH = rFeedKgH) AND ((rFeedKgH - rFeedKgH) = 0.0);
xFinW1 := (rMoistInPct = rMoistInPct) AND ((rMoistInPct - rMoistInPct) = 0.0);
xFinW2 := (rMoistOutPct = rMoistOutPct) AND ((rMoistOutPct - rMoistOutPct) = 0.0);
xFinStm := (rSteamKgH = rSteamKgH) AND ((rSteamKgH - rSteamKgH) = 0.0);
IF (NOT xFinG) OR (NOT xFinW1) OR (NOT xFinW2) OR (NOT xFinStm) THEN
    rWaterAddKgH := 0.0;             // 安全值：加水 0 | safe value, zero water
    rTotalWaterKgH := 0.0;
    rDryMatterKgH := 0.0;
    xReverseMoist := FALSE;
    xValid := FALSE;
    FC_DL_LeafConditioningMoistureCalc := FALSE;
    RETURN;
END_IF

// 段2｜域闸：流量非负、含水率范围、出口不得达 100 %
IF (rFeedKgH < 0.0) OR (rSteamKgH < 0.0)
   OR (rMoistInPct < 0.0) OR (rMoistInPct >= DL_LCM_PCT_MAX)
   OR (rMoistOutPct < 0.0) OR (rMoistOutPct >= DL_LCM_PCT_MAX) THEN
    rWaterAddKgH := 0.0;
    rTotalWaterKgH := 0.0;
    rDryMatterKgH := 0.0;
    xReverseMoist := FALSE;
    xValid := FALSE;
    FC_DL_LeafConditioningMoistureCalc := FALSE;
    RETURN;
END_IF

// 段3｜算法：Gd = G×(100−w1)/100；Wadd = Gd×(w2−w1)/(100−w2)
rDryMatterKgH := rFeedKgH * (DL_LCM_PCT_MAX - rMoistInPct) / DL_LCM_PCT_MAX;
rDenPct := DL_LCM_PCT_MAX - rMoistOutPct;
IF rDenPct > DL_LCM_DEN_MIN THEN
    rWaterAddKgH := rDryMatterKgH * (rMoistOutPct - rMoistInPct) / rDenPct;
ELSE
    rWaterAddKgH := 0.0;             // 理论不可达（段2已排除），防御性兜底 | unreachable defence
END_IF
IF rWaterAddKgH < 0.0 THEN
    xReverseMoist := TRUE;           // 干燥工况：出口按 0 | drying case, zero published
    rWaterAddKgH := 0.0;
ELSE
    xReverseMoist := FALSE;
END_IF

// 段4｜总加水量（蒸汽凝结水按 100 % 计入）
rTotalWaterKgH := rWaterAddKgH + rSteamKgH;
xValid := TRUE;
FC_DL_LeafConditioningMoistureCalc := TRUE;
END_FUNCTION

(* ---- FC_DL_LehrAnnealingScheduleCalc.st ---- *)
(*
  Name: FC_DL_LehrAnnealingScheduleCalc
  Category: DL_Process
  Version: 1.0.0
  Round: R90 / 2026-11-25
  开源溯源：clean-room 自研（族 浮法玻璃锡槽退火，ST 开源生态实测 0 命中，无外部代码引入）
  功能：1) 退火窑温降速率按「区间温差 / 在区间的停留时间」计算：
             停留时间[min] = 区间长度[m] / 线速度[m/min]
             温降速率[°C/min] = (区间进口温度 − 区间出口温度) / 停留时间
           分子方向固定为「进口减出口」：玻璃带沿前进方向降温，故该值为正表示正常降温，
           若为负说明区间在升温（退火窑局部反向，属异常）。速度越快停留时间越短，
           同一温差下温降速率越高，这是本件最核心的方向关系（速度在分母上）。
        2) 与允许退火曲线比较给出 xInSchedule：温降速率必须落在 0 ~ DL_RATE_MAX 的允许带内。
           退火的核心约束是「降温不能过快」，否则玻璃内部产生过大残余应力而炸裂；
           故上限是硬约束，下限 0 用于拦截升温异常。
  边界条件：1) 非有限值闸：四路实值入参统一过 NOT(x > -DL_BIG AND x < DL_BIG)，
           同时拦 NaN 与 Inf，命中即拦断实值通路（fCoolRateCmin 强制 0.0、xInSchedule 强制 FALSE）
           并置无效（R19），无效数据不得判「在曲线上」。
        2) 分母零闸：线速度 ABS > DL_EPS（速度为 0 时停留时间无穷大，温降速率趋于 0，无意义）；
           区间长度 ABS > DL_EPS（长度为 0 时停留时间为 0，温降速率发散）。
        3) 负值闸：区间长度为负、线速度为负判无效（不取绝对值掩盖反向）。
        4) 零值语义：区间温差为 0（等温段）属合法工况，温降速率为 0，判定为在曲线内。
        5) 饱和钳制：温降速率钳 −DL_RATE_MAX ~ +DL_RATE_MAX 的两倍区间，
           防停留时间极小时速率溢出；判定用钳制后的值，保证判据与出口同源。
  量纲自证：停留时间 = m / (m/min) = min；
           fCoolRateCmin = (°C) / min = °C/min，减法两侧同为 °C；
           与 DL_RATE_MAX(°C/min) 同量纲后方可比较，未出现跨量纲混比。
*)

FUNCTION FC_DL_LehrAnnealingScheduleCalc : BOOL
VAR_INPUT
    fZoneInC       : REAL;   // 区间进口玻璃温度 [°C] / Zone inlet glass temperature [°C]
    fZoneOutC      : REAL;   // 区间出口玻璃温度 [°C] / Zone outlet glass temperature [°C]
    fZoneLenM      : REAL;   // 区间长度 [m] / Zone length [m]
    fLineSpeedMmin : REAL;   // 玻璃带线速度 [m/min] / Ribbon line speed [m/min]
END_VAR
VAR_OUTPUT
    fCoolRateCmin  : REAL;   // 温降速率 [°C/min] / Cooling rate [°C/min]
    fResidenceMin  : REAL;   // 区间停留时间（观测用）[min] / Zone residence time [min]
    xInSchedule    : BOOL;   // 在允许退火曲线内 [bool] / Within allowable annealing schedule [bool]
    xValid         : BOOL;   // 计算有效标志 [bool] / Calculation valid flag [bool]
END_VAR
VAR
    _fResidenceRaw : REAL;   // 未饱和的停留时间 [min] / Raw residence time [min]
    _fDeltaTC      : REAL;   // 区间温差（进口 − 出口）[°C] / Zone temperature difference [°C]
    _fRateRaw      : REAL;   // 未饱和的温降速率 [°C/min] / Raw cooling rate [°C/min]
    _fRateClamp    : REAL;   // 饱和钳制后的温降速率 [°C/min] / Clamped cooling rate [°C/min]
END_VAR
VAR CONSTANT
    DL_EPS         : REAL := 1.0E-9;    // 分母零闸阈值 [-] / Division-zero gate threshold [-]
    DL_BIG         : REAL := 1.0E12;    // 非有限值闸量级上限 [-] / Finiteness gate magnitude [-]
    DL_RATE_MAX    : REAL := 15.0;      // 允许温降速率上限 [°C/min] / Allowable cooling rate [°C/min]
    DL_T_HI_C      : REAL := 1200.0;    // 温度量程上限 [°C] / Temperature range high [°C]
END_VAR

(* —— 段 1：非有限值闸（R19：四路入参全覆盖，拦 NaN 与 Inf） —— *)
IF NOT (fZoneInC > -DL_BIG AND fZoneInC < DL_BIG)
   OR NOT (fZoneOutC > -DL_BIG AND fZoneOutC < DL_BIG)
   OR NOT (fZoneLenM > -DL_BIG AND fZoneLenM < DL_BIG)
   OR NOT (fLineSpeedMmin > -DL_BIG AND fLineSpeedMmin < DL_BIG) THEN
    fCoolRateCmin := 0.0;                   // 输出强制 0.0 / Output forced to zero
    fResidenceMin := 0.0;                   // 停留时间强制 0.0 / Residence forced to zero
    xInSchedule := FALSE;                   // 曲线标志强制 FALSE / Schedule flag forced off
    xValid := FALSE;                        // 有效位清零 / Validity cleared
    FC_DL_LehrAnnealingScheduleCalc := FALSE;   // 返回码同源 / Return mirrors validity
    RETURN;                                 // 立即退出 / Immediate exit
END_IF

(* —— 段 2：分母零闸（R4：区间长度与线速度两个分母逐一验证） —— *)
IF (ABS(fZoneLenM) <= DL_EPS) OR (ABS(fLineSpeedMmin) <= DL_EPS) THEN
    fCoolRateCmin := 0.0;                   // 输出强制 0.0 / Output forced to zero
    fResidenceMin := 0.0;                   // 停留时间强制 0.0 / Residence forced to zero
    xInSchedule := FALSE;                   // 曲线标志强制 FALSE / Schedule flag forced off
    xValid := FALSE;                        // 判无效 / Invalid
    FC_DL_LehrAnnealingScheduleCalc := FALSE;   // 返回码同步 / Return synchronised
    RETURN;                                 // 提前退出 / Early exit
END_IF

(* —— 段 3：负值闸（长度与速度为负属组态错误） —— *)
IF (fZoneLenM < 0.0) OR (fLineSpeedMmin < 0.0) THEN
    fCoolRateCmin := 0.0;                   // 输出强制 0.0 / Output forced to zero
    fResidenceMin := 0.0;                   // 停留时间强制 0.0 / Residence forced to zero
    xInSchedule := FALSE;                   // 曲线标志强制 FALSE / Schedule flag forced off
    xValid := FALSE;                        // 判无效 / Invalid
    FC_DL_LehrAnnealingScheduleCalc := FALSE;   // 返回码同步 / Return synchronised
    RETURN;                                 // 提前退出 / Early exit
END_IF

(* —— 段 4：停留时间与温降速率（R22 方向自核：速度在分母，速度快 → 停留短 → 速率高） —— *)
_fResidenceRaw := fZoneLenM / fLineSpeedMmin;                     // 停留时间 [min]
_fDeltaTC := fZoneInC - fZoneOutC;                                // 温差（进口 − 出口）[°C]
_fRateRaw := _fDeltaTC / _fResidenceRaw;                          // 温降速率 [°C/min]

(* —— 段 5：输出单点写盘（出口仅防溢出宽钳，保留真实值；判据另取未夹的原始速率） —— *)
fResidenceMin := LIMIT(0.0, _fResidenceRaw, DL_BIG);              // 停留时间 [min]
_fRateClamp := LIMIT(-DL_BIG, _fRateRaw, DL_BIG);                 // 仅防溢出的宽钳（不夹工艺量程）
fCoolRateCmin := _fRateClamp;                                     // 温降速率出口（真实值，不隐去超速）[°C/min]

(* —— 段 6：有效位单点聚合（温度量程 + 分母为正） —— *)
xValid := (fZoneInC <= DL_T_HI_C) AND (fZoneOutC <= DL_T_HI_C)    // 温度不越量程
          AND (fZoneInC >= 0.0) AND (fZoneOutC >= 0.0)            // 温度非负
          AND (fZoneLenM > DL_EPS)                                // 区间长度为正
          AND (fLineSpeedMmin > DL_EPS);                          // 线速度为正

(* —— 段 7：允许退火曲线判定（0 ~ DL_RATE_MAX 闭区间；负速率即升温，一律判出曲线） —— *)
xInSchedule := xValid AND (_fRateRaw >= 0.0) AND (_fRateRaw <= DL_RATE_MAX);   // 判据用未夹的原始速率，防「钳后判恒真」
FC_DL_LehrAnnealingScheduleCalc := xValid;                        // 返回码：TRUE = 计算可信

END_FUNCTION

(* ---- FC_DL_LifterCycleTimeEst.st ---- *)
(*
  ============================================================
  组件名 : FC_DL_LifterCycleTimeEst
  分类   : DL_Process
  功能   : 提升机单循环节拍估算，由层高与层数求往复升降时间并叠加开关门与货叉时间
  复杂度 : C1
  版本   : 1.0.0
  作者   : 道莅工业代码库工厂 / R81
  日期   : 2026-11-24
  开源溯源 : clean-room（no upstream）—— 依据公开工程公式自研，未复制任何上游实现
  红线自检 : R1 无GVL/R2 无物理地址/R3 纯IEC/R4 防除零/R5 双语注释
  接口说明 :
      单循环 = 2*(层高*(层数-1)/提升速度) + 2*开关门时间 + 2*货叉时间，即一取一放完整往复。
      层数要求 >= 2，层数 1 时无层间位移，节拍模型不成立，直接判无效。
      rCap 由 3600/rCycle 折算，rCycle 非正时不做除法，仅保留时间输出并判无效。
  ============================================================
*)
FUNCTION FC_DL_LifterCycleTimeEst : BOOL
VAR_INPUT
    bEnable   : BOOL; // 使能：TRUE 时计算 / Enable: TRUE to compute
    bErr      : BOOL; // 外部故障：TRUE 时立即退出并置结果无效 / External fault: TRUE aborts with invalid result
    rLiftH    : REAL; // 层间高度 [m] / height between two adjacent levels [m]
    iLayers   : INT;  // 货架总层数 [层] / total number of levels [level]
    rVlift    : REAL; // 提升额定速度 [m/s] / rated lifting speed [metre per second]
    rTdoor    : REAL; // 单次开关门时间 [s] / door open close time for one operation [s]
    rTfork    : REAL; // 单次货叉伸缩时间 [s] / fork extend retract time for one operation [s]
END_VAR
VAR_OUTPUT
    rCycle_s  : REAL; // 单循环节拍时间 [s] / single cycle time [s]
    rCap      : REAL; // 折算产能 [件/小时] / equivalent capacity [piece per hour]
    bValid    : BOOL; // 输出有效：TRUE 表示结果可用 / Output valid
END_VAR
VAR CONSTANT
    DL_R_MAX   : REAL := 3.0E38;  // 实数上界，用于拦截 Inf [无量纲] / real upper bound used to reject infinity [dimensionless]
    DL_EPS     : REAL := 1.0E-12; // 除零判定阈值 [无量纲] / division guard threshold [dimensionless]
    DL_SEC_H   : REAL := 3600.0;  // 每小时秒数 [s/h] / seconds per hour [second per hour]
    DL_TWO     : REAL := 2.0;     // 往复行程倍数 [无量纲] / round trip multiplier [dimensionless]
END_VAR
VAR
    _bFin    : BOOL := FALSE; // 输入有限性判定汇总 / aggregated finiteness verdict of the inputs
    _rTravel : REAL := 0.0;   // 单程升降时间 [s] / one way travel time [s]
    _rLayers : REAL := 0.0;   // 层数折算实数 [无量纲] / level count cast to real [dimensionless]
END_VAR

    // 段 1｜出口预置
    rCycle_s := 0.0;
    rCap := 0.0;
    bValid := FALSE;
    // 段 2｜使能闸与外部故障闸
    IF NOT bEnable THEN
        RETURN;
    END_IF;
    IF bErr THEN
        RETURN;
    END_IF;
    // 段 3｜非有限闸
    _bFin := (rLiftH = rLiftH) AND (ABS(rLiftH) <= DL_R_MAX) AND (rVlift = rVlift) AND (ABS(rVlift) <= DL_R_MAX) AND (rTdoor = rTdoor) AND (ABS(rTdoor) <= DL_R_MAX) AND (rTfork = rTfork) AND (ABS(rTfork) <= DL_R_MAX);
    IF NOT _bFin THEN
        RETURN;
    END_IF;
    // 段 4｜域闸：速度必须严格为正，层数必须 >= 2，时间与层高不得为负
    IF ABS(rVlift) <= DL_EPS THEN
        RETURN;
    END_IF;
    IF iLayers < 2 THEN
        RETURN;
    END_IF;
    IF (rLiftH < 0.0) OR (rVlift < 0.0) OR (rTdoor < 0.0) OR (rTfork < 0.0) THEN
        RETURN;
    END_IF;
    // 段 5｜单程升降时间：层数减一得到层间跨距个数
    _rLayers := INT_TO_REAL(iLayers);
    _rTravel := rLiftH * (_rLayers - 1.0) / rVlift;
    // 段 6｜单循环时间：升降往复加两次开关门加两次货叉
    rCycle_s := DL_TWO * _rTravel + DL_TWO * rTdoor + DL_TWO * rTfork;
    // 段 7｜产能折算：必须再次确认周期严格为正才允许做除法
    IF rCycle_s > DL_EPS THEN
        rCap := DL_SEC_H / rCycle_s;
    ELSE
        rCap := 0.0;
        bValid := FALSE;
        FC_DL_LifterCycleTimeEst := bValid;
        RETURN;
    END_IF;
    bValid := TRUE;
    FC_DL_LifterCycleTimeEst := bValid;
END_FUNCTION

(* ---- FC_DL_LyoChamberLeakRateCalc.st ---- *)
(*
  Name: FC_DL_LyoChamberLeakRateCalc
  Category: DL_Process
  Version: 1.0.0
  Round: R91 / 2026-11-25
  开源溯源：clean-room 自研（族 制药冻干真空冷冻干燥，ST 开源生态实测 0 命中，无外部代码引入）
  功能：1) 腔体泄漏率按压力升试验法（pressure rise test）计算：
           Q = dP * V / t，dP 为隔离后腔内压力升幅 [mbar]、V 为腔体内容积 [L]、t 为测试时长 [s]，
           结果单位 mbar*L/s，是冻干机 GMP 验证的法定泄漏率指标。
        2) 合格判据：Q <= fLeakMaxMbarLs 输出 xPass；同时给出负荷率 fLeakLoadPct = Q / 上限 * 100，
           便于观察密封状态的趋势劣化（负荷率单调上升意味着门封老化）。
        3) 压力升幅方向校验：升幅必须 > 0（隔离后压力只能升，若为负说明隔离阀未关严或
           仍有抽气，测试无效），负升幅判 xValid = FALSE 而非取绝对值。
  边界条件：1) 非有限值闸：四路实值入参先过 NOT(x > -DL_BIG AND x < DL_BIG)，同时拦 NaN 与 Inf，
           命中即闸断实值通路（泄漏率与负荷率强制 0.0），不得只置标志（R19）。
        2) 时间零闸：测试时长 fTestTimeS 必须 > DL_EPS（泄漏率式分母），
           否则判无效并清零，不得输出无穷大泄漏率。
        3) 容积零闸：腔体容积 fVolumeL 必须 > DL_EPS（乘子为零会使一切泄漏率归零，
           把「未接容积组态」伪装成「密封完好」）。
        4) 判据取原始值（R24）：合格判定使用钳制前的 _fLeakRaw，不得先钳再判。
        5) 物理域钳制：泄漏率钳 0.0 ~ DL_LEAK_HI；负荷率钳 0.0 ~ DL_PCT_HI。
        6) 纯函数无状态：本件只算一次测试结果，多次测试的平均与趋势判断由上层质量模块承担。
  量纲自证：Q = (mbar)*(L)/(s) = mbar*L/s，三个因子量纲直乘/直除，无跨量纲混算；
           fLeakLoadPct = (mbar*L/s)/(mbar*L/s)*100 = 无因次百分数 [%]，量纲合法。
  修订历史 Revision :
    2026-11-25  v1.0.0  R91 首版
*)

FUNCTION FC_DL_LyoChamberLeakRateCalc : BOOL
VAR_INPUT
    fPressRiseMbar   : REAL;   // 测试期腔内压力升幅 [mbar] / Chamber pressure rise during the test [mbar]
    fVolumeL         : REAL;   // 腔体（含管路）内容积 [L] / Chamber and piping internal volume [L]
    fTestTimeS       : REAL;   // 测试时长 [s] / Test duration [s]
    fLeakMaxMbarLs   : REAL;   // 泄漏率合格上限 [mbar*L/s] / Leak rate acceptance limit [mbar*L/s]
END_VAR
VAR_OUTPUT
    fLeakRateMbarLs  : REAL;   // 实测泄漏率 [mbar*L/s] / Measured leak rate [mbar*L/s]
    fLeakLoadPct     : REAL;   // 泄漏率对合格上限的负荷率 [%] / Leak load ratio against the limit [%]
    xPass            : BOOL;   // 合格标志 [bool] / Acceptance flag [bool]
    xValid           : BOOL;   // 计算有效标志 [bool] / Calculation valid flag [bool]
END_VAR
VAR
    _fLeakRaw        : REAL;   // 钳制前的原始泄漏率 [mbar*L/s] / Raw leak rate before limiting [mbar*L/s]
    _fLoadRawPct     : REAL;   // 钳制前的原始负荷率 [%] / Raw load ratio before limiting [%]
END_VAR
VAR CONSTANT
    DL_EPS           : REAL := 1.0E-9;    // 数值零闸阈值 [-] / Numeric zero gate threshold [-]
    DL_BIG           : REAL := 1.0E12;    // 非有限值闸量级上限 [-] / Finiteness gate magnitude [-]
    DL_PCT           : REAL := 100.0;     // 百分比换算因子 [%] / Percent conversion factor [%]
    DL_PCT_HI        : REAL := 1000.0;    // 负荷率显示上限（允许超 100 % 报警）[%] / Load ratio display ceiling [%]
    DL_LEAK_HI       : REAL := 100.0;     // 泄漏率物理上限 [mbar*L/s] / Leak rate physical upper bound [mbar*L/s]
END_VAR

(* —— 段 1：非有限值闸（R19：闸断实值通路） —— *)
IF NOT (fPressRiseMbar > -DL_BIG AND fPressRiseMbar < DL_BIG)
   OR NOT (fVolumeL > -DL_BIG AND fVolumeL < DL_BIG)
   OR NOT (fTestTimeS > -DL_BIG AND fTestTimeS < DL_BIG)
   OR NOT (fLeakMaxMbarLs > -DL_BIG AND fLeakMaxMbarLs < DL_BIG) THEN
    fLeakRateMbarLs := 0.0;                 // 输出强制 0.0，切断污染源 / Force zero, cut polluted path
    fLeakLoadPct := 0.0;                    // 负荷率强制 0.0 / Load ratio forced to zero
    xPass := FALSE;                         // 失效侧不得判合格（安全侧）/ Must not report pass when invalid
    xValid := FALSE;                        // 有效位清零 / Validity cleared
    FC_DL_LyoChamberLeakRateCalc := FALSE;  // 返回码与有效位同源 / Return mirrors validity
    RETURN;                                 // 立即退出 / Immediate exit
END_IF

(* —— 段 2：时间零闸与参数域闸（时间式为分母，容积为乘子都须为正） —— *)
IF (fTestTimeS <= DL_EPS)                                         // 测试时长不可为零
   OR (fVolumeL <= DL_EPS)                                        // 容积不可为零（防「未组态」伪装成完好）
   OR (fLeakMaxMbarLs <= DL_EPS) THEN                             // 合格上限必须已组态
    fLeakRateMbarLs := 0.0;                 // 参数不可用即无泄漏率 / No parameter, no leak rate
    fLeakLoadPct := 0.0;                    // 负荷率不可算 / Load ratio not computable
    xPass := FALSE;                         // 判不合格 / Not accepted
    xValid := FALSE;                        // 判无效 / Invalid
    FC_DL_LyoChamberLeakRateCalc := FALSE;  // 返回码同步 / Return synchronised
    RETURN;                                 // 提前退出 / Early exit
END_IF

(* —— 段 3：主算式（不钳制，先出原始值供段 4 判据使用，R24） —— *)
_fLeakRaw := fPressRiseMbar * fVolumeL / fTestTimeS;                              // 泄漏率 [mbar*L/s]
_fLoadRawPct := _fLeakRaw / fLeakMaxMbarLs * DL_PCT;                              // 负荷率 [%]

(* —— 段 4：判据（取原始值；单点 BOOL 聚合避免多处赋 FALSE 覆盖） —— *)
xValid := (fPressRiseMbar > 0.0)                                                  // 升幅必须为正（隔离有效性）
          AND (_fLeakRaw >= 0.0)                                                  // 泄漏率不得为负
          AND (_fLeakRaw <= DL_LEAK_HI)                                           // 不得超物理上限（量级异常）
          AND (fLeakMaxMbarLs <= DL_LEAK_HI);                                     // 合格上限须在物理域内
xPass := (_fLeakRaw <= fLeakMaxMbarLs) AND xValid;                                // 不越上限且计算可信才判合格

(* —— 段 5：输出单点写盘（钳制到物理域内，判定结果已在段 4 定案） —— *)
fLeakRateMbarLs := LIMIT(0.0, _fLeakRaw, DL_LEAK_HI);                             // 泄漏率钳 0..物理上限
fLeakLoadPct := LIMIT(0.0, _fLoadRawPct, DL_PCT_HI);                              // 负荷率钳 0..显示上限 [%]
FC_DL_LyoChamberLeakRateCalc := xValid;                                           // 返回码：TRUE = 计算可信

END_FUNCTION
